(* IEC 61131-3 sources: PLC-IsaVODE/PLC-IsaVODE/samples/plc-programs (part 14) *)

(* ---- 100-RES_NTC.ST ---- *)
FUNCTION RES_NTC:REAL

	VAR_INPUT
		T :	REAL;
		RN :	REAL;
		B :	REAL;
	END_VAR

	RES_NTC := RN * EXP(B * (1.0 / (T+273.15) - 0.00335401643468053));

END_FUNCTION

PROGRAM program0

	VAR
		T :	REAL;
		RN :	REAL;
		B :	REAL;

		OUT :	REAL;
	END_VAR
		OUT := RES_NTC(T, RN, B);

END_PROGRAM

CONFIGURATION Config0

	RESOURCE Res0 ON PLC
		TASK task0(INTERVAL := T#20ms,PRIORITY := 0);
		PROGRAM instance0 WITH task0 : program0;
	END_RESOURCE

END_CONFIGURATION

(* ---- 101-WINDOW2.ST ---- *)
FUNCTION WINDOW2:BOOL
	VAR_INPUT
		LOW :	REAL;
		IN :	REAL;
		HIGH :	REAL;
	END_VAR
	window2 := (in <= high) AND (in >= low);
END_FUNCTION

PROGRAM program0
  	VAR
		LOW :	REAL;
		IN :	REAL;
		HIGH :	REAL;
		CEIL5_OUT : BOOL;
	END_VAR

  	CEIL5_OUT := window2(LOW, IN, HIGH);
END_PROGRAM

CONFIGURATION Config0
  	RESOURCE Res0 ON PLC
    	TASK task0(INTERVAL := T#20ms,PRIORITY := 0);
    	PROGRAM instance0 WITH task0 : program0;
  	END_RESOURCE
END_CONFIGURATION

(* ---- 102-F_LIN.ST ---- *)
FUNCTION F_LIN:REAL
	VAR_INPUT
		X :	REAL;
		A :	REAL;
		B :	REAL;
	END_VAR

	F_lin := A * X + B;
END_FUNCTION

PROGRAM program0
  VAR
    LocalVar0 : REAL;
	LocalVar1 : REAL;
	LocalVar2 : REAL;
	  LocalOUT  : REAL;
  END_VAR
  	LocalOUT := F_LIN(LocalVar0, LocalVar1, LocalVar2);
END_PROGRAM

CONFIGURATION Config0
  RESOURCE Res0 ON PLC
    TASK task0(INTERVAL := T#20ms,PRIORITY := 0);
    PROGRAM instance0 WITH task0 : program0;
  END_RESOURCE
END_CONFIGURATION

(* ---- 103-TN_SC_SHADOW_ATTR.ST ---- *)
FUNCTION TN_SC_SHADOW_ATTR:BYTE

	VAR_INPUT
		Iby_ATTR :	BYTE;
	END_VAR

	TN_SC_SHADOW_ATTR := ((Iby_ATTR AND BYTE#2#11110000) OR BYTE#2#00001000);

END_FUNCTION

PROGRAM program0
	VAR
		Iby_ATTR :	BYTE;
		CEIL5_OUT : BYTE;
	END_VAR

  	CEIL5_OUT := TN_SC_SHADOW_ATTR(Iby_ATTR);
END_PROGRAM

CONFIGURATION Config0

  RESOURCE Res0 ON PLC
    TASK task0(INTERVAL := T#20ms,PRIORITY := 0);
    PROGRAM instance0 WITH task0 : program0;
  END_RESOURCE
END_CONFIGURATION

(* ---- 104-DEC1.ST ---- *)
FUNCTION DEC1:INT

	VAR_INPUT
		X :	INT;
		N :	INT;
	END_VAR

	IF X = 0 THEN
		DEC1 := N - 1;
	ELSE
		DEC1 := X - 1;
	END_IF;

END_FUNCTION

PROGRAM program0
  VAR
    LocalVar0 : INT;
	LocalVar1 : INT;
	LocalOUT  : INT;
  END_VAR
  	LocalOUT := DEC1(LocalVar0, LocalVar1);
END_PROGRAM

CONFIGURATION Config0
  RESOURCE Res0 ON PLC
    TASK task0(INTERVAL := T#20ms,PRIORITY := 0);
    PROGRAM instance0 WITH task0 : program0;
  END_RESOURCE
END_CONFIGURATION

(* ---- 105-INC.ST ---- *)
FUNCTION INC:INT
	VAR_INPUT
		X :	INT;
		D :	INT;
		M :	INT;
	END_VAR

	inc := (X + D + M + 1) MOD (M + 1);
END_FUNCTION

PROGRAM program0
  VAR
    LocalVar0 : INT;
	LocalVar1 : INT;
	LocalVar2 : INT;
	LocalOUT  : INT;
  END_VAR
  	LocalOUT := INC(LocalVar0, LocalVar1,LocalVar2);
END_PROGRAM

CONFIGURATION Config0
  RESOURCE Res0 ON PLC
    TASK task0(INTERVAL := T#20ms,PRIORITY := 0);
    PROGRAM instance0 WITH task0 : program0;
  END_RESOURCE
END_CONFIGURATION

(* ---- 106-BIT_TOGGLE_B.ST ---- *)
FUNCTION BIT_TOGGLE_B:BYTE
	VAR_INPUT
		IN :	BYTE;
		POS :	INT;
	END_VAR

	BIT_TOGGLE_B := SHL(BYTE#1, POS) XOR IN;
END_FUNCTION

PROGRAM program0
  VAR
    LocalVar0 : BYTE;
    LocalVar1 : INT;
    CEIL5_OUT : BYTE;
  END_VAR

  CEIL5_OUT := BIT_TOGGLE_B(LocalVar0, LocalVar1);
END_PROGRAM

CONFIGURATION Config0

  RESOURCE Res0 ON PLC
    TASK task0(INTERVAL := T#20ms,PRIORITY := 0);
    PROGRAM instance0 WITH task0 : program0;
  END_RESOURCE
END_CONFIGURATION

(* ---- 107-BIT_TOGGLE_W.ST ---- *)
FUNCTION BIT_TOGGLE_W:WORD
	VAR_INPUT
		IN :	WORD;
		POS :	INT;
	END_VAR

	BIT_TOGGLE_W := SHL(WORD#1, POS) XOR IN;
END_FUNCTION

PROGRAM program0
  VAR
    LocalVar0 : WORD;
    LocalVar1 : INT;
    CEIL5_OUT : WORD;
  END_VAR

  CEIL5_OUT := BIT_TOGGLE_W(LocalVar0, LocalVar1);
END_PROGRAM

CONFIGURATION Config0

  RESOURCE Res0 ON PLC
    TASK task0(INTERVAL := T#20ms,PRIORITY := 0);
    PROGRAM instance0 WITH task0 : program0;
  END_RESOURCE
END_CONFIGURATION

(* ---- 108-RES_NI.ST ---- *)
FUNCTION RES_NI:REAL

	VAR_INPUT
		T :	REAL;
		R0 :	REAL;
	END_VAR

	VAR
		T2 :	REAL;
	END_VAR

	T2 := T*T;
	Res_NI := R0 + 0.5485*T + 0.665E-3*T2 + 2.805E-9*T2*T2;

END_FUNCTION

PROGRAM program0

	VAR
		T :	REAL;
		R0 :	REAL;

		OUT :	REAL;
	END_VAR
	OUT := RES_NI(T, R0);

END_PROGRAM

CONFIGURATION Config0

	RESOURCE Res0 ON PLC
		TASK task0(INTERVAL := T#20ms,PRIORITY := 0);
		PROGRAM instance0 WITH task0 : program0;
	END_RESOURCE

END_CONFIGURATION

(* ---- 109-TANK_VOL2.ST ---- *)
FUNCTION TANK_VOL2:REAL

	VAR_INPUT
		TR :	REAL;
		H :	REAL;
	END_VAR

	TANK_VOL2 := 3.14159265358979323846264338327950288 * H * H * (TR - H / 3.0);

END_FUNCTION

PROGRAM program0
  VAR
    TR :	REAL;
	H :	REAL;
    CEIL5_OUT : REAL;
  END_VAR

  CEIL5_OUT := TANK_VOL2(TR, H);
END_PROGRAM

CONFIGURATION Config0

  RESOURCE Res0 ON PLC
    TASK task0(INTERVAL := T#20ms,PRIORITY := 0);
    PROGRAM instance0 WITH task0 : program0;
  END_RESOURCE
END_CONFIGURATION

(* ---- 11-SWAP_BYTE.ST ---- *)
FUNCTION SWAP_BYTE:WORD

	VAR_INPUT
		IN :	WORD;
	END_VAR

	Swap_Byte := ROL(in,8);

END_FUNCTION

PROGRAM program0

	VAR
		IN :	WORD;
		CEIL5_OUT : WORD;
	END_VAR

	CEIL5_OUT := SWAP_BYTE(IN);

END_PROGRAM

CONFIGURATION Config0

	RESOURCE Res0 ON PLC
		TASK task0(INTERVAL := T#20ms,PRIORITY := 0);
		PROGRAM instance0 WITH task0 : program0;
	END_RESOURCE

END_CONFIGURATION

(* ---- 110-YEAR_END.ST ---- *)
FUNCTION YEAR_END:UDINT

	VAR_INPUT
		Y :	INT;
	END_VAR

	YEAR_END := DWORD_TO_UDINT(SHR(UDINT_TO_DWORD(INT_TO_UDINT(y) * UDINT#1461 - UDINT#2876712), 2)) * UDINT#86400;

END_FUNCTION

PROGRAM program0
  VAR
    Y : INT;
    CEIL5_OUT : UDINT;
  END_VAR

  CEIL5_OUT := YEAR_END(Y);
END_PROGRAM

CONFIGURATION Config0

  RESOURCE Res0 ON PLC
    TASK task0(INTERVAL := T#20ms,PRIORITY := 0);
    PROGRAM instance0 WITH task0 : program0;
  END_RESOURCE
END_CONFIGURATION

(* ---- 111-IP4_CHECK.ST ---- *)
FUNCTION IP4_CHECK:BOOL

	VAR_INPUT
		NIP :	DWORD;
		LIP :	DWORD;
		SM :	DWORD;
	END_VAR

	IP4_CHECK := (NIP AND sm) = (LIP AND SM);

END_FUNCTION

PROGRAM program0
	VAR
		NIP :	DWORD;
		LIP :	DWORD;
		SM :	DWORD;
		CEIL5_OUT : BOOL;
	END_VAR

  	CEIL5_OUT := IP4_CHECK(NIP, LIP, SM);
END_PROGRAM

CONFIGURATION Config0

  RESOURCE Res0 ON PLC
    TASK task0(INTERVAL := T#20ms,PRIORITY := 0);
    PROGRAM instance0 WITH task0 : program0;
  END_RESOURCE
END_CONFIGURATION

(* ---- 112-ELLIPSE_A.ST ---- *)
FUNCTION ELLIPSE_A:REAL
	VAR_INPUT
		R1 :	REAL;
		R2 :	REAL;
	END_VAR

	ellipse_A := 3.14159265358979323846264338327950288 * R1 * R2;

END_FUNCTION

PROGRAM program0
  VAR
    LocalVar0 : REAL;
	LocalVar1 : REAL;
	  LocalOUT  : REAL;
  END_VAR
  	LocalOUT := ELLIPSE_A(LocalVar0, LocalVar1);
END_PROGRAM

CONFIGURATION Config0
  RESOURCE Res0 ON PLC
    TASK task0(INTERVAL := T#20ms,PRIORITY := 0);
    PROGRAM instance0 WITH task0 : program0;
  END_RESOURCE
END_CONFIGURATION

(* ---- 113-F_POWER.ST ---- *)
FUNCTION F_POWER:REAL
	VAR_INPUT
		A :	REAL;
		X :	REAL;
		N :	REAL;
	END_VAR

	f_power := a * EXPT(X,N);
END_FUNCTION

PROGRAM program0
  VAR
    LocalVar0 : REAL;
	LocalVar1 : REAL;
	LocalVar2 : REAL;
	  LocalOUT  : REAL;
  END_VAR
  	LocalOUT := F_POWER(LocalVar0, LocalVar1, LocalVar2);
END_PROGRAM

CONFIGURATION Config0
  RESOURCE Res0 ON PLC
    TASK task0(INTERVAL := T#20ms,PRIORITY := 0);
    PROGRAM instance0 WITH task0 : program0;
  END_RESOURCE
END_CONFIGURATION

(* ---- 114-TANH.ST ---- *)
FUNCTION TANH:REAL

	VAR_INPUT
		X :	REAL;
	END_VAR

	IF X > 20.0 THEN
		TANH := 1.0;
	ELSIF X < -20.0 THEN
		TANH := -1.0;
	ELSE
		TANH := 1.0 - 2.0 / (EXP(2.0 * x) + 1.0);
	END_IF;

END_FUNCTION

PROGRAM program0

	VAR
		X :	REAL;
		CEIL5_OUT : REAL;
	END_VAR

	CEIL5_OUT := TANH(X);

END_PROGRAM

CONFIGURATION Config0

	RESOURCE Res0 ON PLC
		TASK task0(INTERVAL := T#20ms,PRIORITY := 0);
		PROGRAM instance0 WITH task0 : program0;
	END_RESOURCE

END_CONFIGURATION

(* ---- 115-BIT_TOGGLE_DW.ST ---- *)
FUNCTION BIT_TOGGLE_DW:DWORD
	VAR_INPUT
		IN :	DWORD;
		POS :	INT;
	END_VAR

	BIT_TOGGLE_DW := SHL(DWORD#1, POS) XOR IN;

END_FUNCTION

PROGRAM program0
  VAR
    LocalVar0 : DWORD;
    LocalVar1 : INT;
    CEIL5_OUT : DWORD;
  END_VAR

  CEIL5_OUT := BIT_TOGGLE_DW(LocalVar0, LocalVar1);
END_PROGRAM

CONFIGURATION Config0

  RESOURCE Res0 ON PLC
    TASK task0(INTERVAL := T#20ms,PRIORITY := 0);
    PROGRAM instance0 WITH task0 : program0;
  END_RESOURCE
END_CONFIGURATION

(* ---- 116-SIGMOID.ST ---- *)
FUNCTION SIGMOID:REAL

	VAR_INPUT
		X :	REAL;
	END_VAR

	IF X > 20.0 THEN
		SIGMOID := 1.0;
	ELSIF x < -85.0 THEN
		SIGMOID := 0.0;
	ELSE
		SIGMOID := 1.0 / (1.0 + EXP(-X));
	END_IF;

END_FUNCTION

PROGRAM program0

	VAR
		X :	REAL;
		CEIL5_OUT : REAL;
	END_VAR

	CEIL5_OUT := SIGMOID(X);

END_PROGRAM

CONFIGURATION Config0

	RESOURCE Res0 ON PLC
		TASK task0(INTERVAL := T#20ms,PRIORITY := 0);
		PROGRAM instance0 WITH task0 : program0;
	END_RESOURCE

END_CONFIGURATION

(* ---- 117-LEAP_OF_DATE.ST ---- *)
FUNCTION LEAP_OF_DATE:BOOL

	VAR_INPUT
		IDATE :	UDINT;
	END_VAR

	LEAP_OF_DATE := SHL(UDINT_TO_DWORD((idate + UDINT#43200) / UDINT#31557600), 30) = DWORD#16#80000000;

END_FUNCTION

PROGRAM program0
  VAR
    LocalVar0 : UDINT;
	LocalOUT  : BOOL;
  END_VAR
  	LocalOUT := LEAP_OF_DATE(LocalVar0);
END_PROGRAM

CONFIGURATION Config0
  RESOURCE Res0 ON PLC
    TASK task0(INTERVAL := T#20ms,PRIORITY := 0);
    PROGRAM instance0 WITH task0 : program0;
  END_RESOURCE
END_CONFIGURATION

(* ---- 118-DIFFER.ST ---- *)
FUNCTION DIFFER:BOOL
	VAR_INPUT
		IN1 :	REAL;
		IN2 :	REAL;
		X :	REAL;
	END_VAR

	DIFFER := ABS(in1 - in2) > X;
END_FUNCTION

PROGRAM program0
  VAR
    LocalVar0 : REAL;
	LocalVar1 : REAL;
	LocalVar2 : REAL;
	LocalOUT  : BOOL;
  END_VAR
  	LocalOUT := DIFFER(LocalVar0, LocalVar1, LocalVar2);
END_PROGRAM

CONFIGURATION Config0
  RESOURCE Res0 ON PLC
    TASK task0(INTERVAL := T#20ms,PRIORITY := 0);
    PROGRAM instance0 WITH task0 : program0;
  END_RESOURCE
END_CONFIGURATION

(* ---- 119-DEAD_ZONE.ST ---- *)
FUNCTION DEAD_ZONE:REAL

	VAR_INPUT
		X :	REAL;
		L :	REAL;
	END_VAR

	IF ABS(x) > L THEN
		dead_zone := X;
	ELSE
		DEAD_ZONE := 0.0;
	END_IF;

END_FUNCTION

PROGRAM program0
  VAR
    LocalVar0 : REAL;
	LocalVar1 : REAL;
	LocalOUT  : REAL;
  END_VAR
  	LocalOUT := DEAD_ZONE(LocalVar0, LocalVar1);
END_PROGRAM

CONFIGURATION Config0
  RESOURCE Res0 ON PLC
    TASK task0(INTERVAL := T#20ms,PRIORITY := 0);
    PROGRAM instance0 WITH task0 : program0;
  END_RESOURCE
END_CONFIGURATION

(* ---- 12-ISC_CTRL.ST ---- *)
FUNCTION ISC_CTRL:BOOL

	VAR_INPUT
		IN :	BYTE;
	END_VAR

	ISC_CTRL := IN < BYTE#32 OR IN = BYTE#127;

END_FUNCTION

PROGRAM program0
	VAR
		IN : BYTE;
		OUT : BOOL;
	END_VAR

	OUT := ISC_CTRL(IN);
END_PROGRAM

CONFIGURATION Config0

	RESOURCE Res0 ON PLC
		TASK task0(INTERVAL := T#20ms,PRIORITY := 0);
		PROGRAM instance0 WITH task0 : program0;
	END_RESOURCE

END_CONFIGURATION

(* ---- 120-SQRTN.ST ---- *)
FUNCTION SQRTN:REAL

	VAR_INPUT
		X :	REAL;
		N :	INT;
	END_VAR

	IF N > 0 THEN
		SQRTN := EXP(LN(x) / INT_TO_REAL(n));
	ELSE
		SQRTN := 0.0;
	END_IF;

END_FUNCTION

PROGRAM program0
	VAR
		LocalVar0 : REAL;
		LocalVar1 : INT;
		LocalOUT  : REAL;
	END_VAR

 	LocalOUT := SQRTN(LocalVar0, LocalVar1);

END_PROGRAM

CONFIGURATION Config0

	RESOURCE Res0 ON PLC
		TASK task0(INTERVAL := T#20ms,PRIORITY := 0);
		PROGRAM instance0 WITH task0 : program0;
	END_RESOURCE

END_CONFIGURATION

(* ---- 122-DWORD_OF_WORD.ST ---- *)
FUNCTION DWORD_OF_WORD:DWORD

	VAR_INPUT
		W1 :	WORD;
		W0 :	WORD;
	END_VAR

	DWORD_OF_WORD := SHL(WORD_TO_DWORD(W1),16) OR WORD_TO_DWORD(W0);

END_FUNCTION

PROGRAM program0
  VAR
    LocalVar0 : WORD;
	LocalVar1 : WORD;
	LocalOUT  : DWORD;
  END_VAR
  	LocalOUT := DWORD_OF_WORD(LocalVar0, LocalVar1);
END_PROGRAM

CONFIGURATION Config0
  RESOURCE Res0 ON PLC
    TASK task0(INTERVAL := T#20ms,PRIORITY := 0);
    PROGRAM instance0 WITH task0 : program0;
  END_RESOURCE
END_CONFIGURATION

(* ---- 123-WCT.ST ---- *)
FUNCTION WCT:REAL

	VAR_INPUT
		T :	REAL;
		V :	REAL;
	END_VAR

	IF V < 5.0 OR T > 10.0 THEN
		WCT := T;
	ELSE
		WCT := 13.12 + 0.6215 * T +(0.3965 * T - 11.37) * EXP(LN(v) * 0.16);
	END_IF;

END_FUNCTION

PROGRAM program0
	VAR
		T :	REAL;
		V :	REAL;
		CEIL5_OUT : REAL;
	END_VAR

  	CEIL5_OUT := WCT(T, V);
END_PROGRAM

CONFIGURATION Config0

  RESOURCE Res0 ON PLC
    TASK task0(INTERVAL := T#20ms,PRIORITY := 0);
    PROGRAM instance0 WITH task0 : program0;
  END_RESOURCE
END_CONFIGURATION

(* ---- 124-TEMP_NTC.ST ---- *)
FUNCTION TEMP_NTC:REAL

VAR_INPUT
	RES :	REAL;
	RN :	REAL;
	B :	REAL;
END_VAR

IF res > 0.0 THEN
	TEMP_NTC := B * 298.15 / (B + LN(RES / RN) * 298.15) -273.15;
END_IF;

END_FUNCTION

PROGRAM program0
  	VAR
		RES :	REAL;
		RN :	REAL;
		B :	REAL;
    	CEIL5_OUT : REAL;
  	END_VAR

  	CEIL5_OUT := TEMP_NTC(RES, RN, B);
END_PROGRAM

CONFIGURATION Config0
	RESOURCE Res0 ON PLC
		TASK task0(INTERVAL := T#20ms,PRIORITY := 0);
		PROGRAM instance0 WITH task0 : program0;
	END_RESOURCE
END_CONFIGURATION

(* ---- 125-SCALE.ST ---- *)
FUNCTION SCALE:REAL

	VAR_INPUT
		X :	REAL;
		K :	REAL;
		O :	REAL;
		MX :	REAL;
		MN :	REAL;
	END_VAR

	SCALE := LIMIT(MN, X * K + O, MX);

END_FUNCTION

PROGRAM program0
  VAR
    X :	REAL;
	K :	REAL;
	O :	REAL;
	MX :	REAL;
	MN :	REAL;
    CEIL5_OUT : REAL;
  END_VAR

  CEIL5_OUT := SCALE(X, K, O, MX, MN);
END_PROGRAM

CONFIGURATION Config0

  RESOURCE Res0 ON PLC
    TASK task0(INTERVAL := T#20ms,PRIORITY := 0);
    PROGRAM instance0 WITH task0 : program0;
  END_RESOURCE
END_CONFIGURATION

(* ---- 126-_MOD_INT.ST ---- *)
FUNCTION _MOD_INT:INT
  VAR_INPUT
    IN :	INT;
    DIVISOR :	INT;
  END_VAR

  IF IN = 0 THEN
    _MOD_INT := 0;
  ELSE
    _MOD_INT := IN MOD DIVISOR;
  END_IF;
END_FUNCTION

PROGRAM program0
  VAR
    LocalVar0 : INT;
    LocalVar1 : INT;
	  LocalOUT  : INT;
  END_VAR

  LocalOUT := _MOD_INT(LocalVar0, LocalVar1);
END_PROGRAM

CONFIGURATION Config0
  RESOURCE Res0 ON PLC
    TASK task0(INTERVAL := T#20ms,PRIORITY := 0);
    PROGRAM instance0 WITH task0 : program0;
  END_RESOURCE
END_CONFIGURATION

(* ---- 127-INC2.ST ---- *)
FUNCTION INC2:INT

	VAR_INPUT
		X :	INT;
		D :	INT;
		L :	INT;
		U :	INT;
	END_VAR

	VAR
		tmp :	INT;
	END_VAR

	tmp := U - L + 1;
	INC2 := (X + D - L + tmp) MOD tmp + L;

END_FUNCTION

PROGRAM program0
	VAR
		X :	INT;
		D :	INT;
		L :	INT;
		U :	INT;
		CEIL5_OUT : INT;
	END_VAR

  	CEIL5_OUT := INC2(X, D, L, U);
END_PROGRAM

CONFIGURATION Config0

	RESOURCE Res0 ON PLC
		TASK task0(INTERVAL := T#20ms,PRIORITY := 0);
		PROGRAM instance0 WITH task0 : program0;
	END_RESOURCE

END_CONFIGURATION

(* ---- 128-TEMP_SI.ST ---- *)
FUNCTION TEMP_SI:REAL
	VAR_INPUT
		RES :	REAL;
		VAR_RS:	REAL;
		TS :	REAL;
	END_VAR

	TEMP_SI := (-7.64E-3 + SQRT(RES/VAR_RS* 6.64E-5 - 0.803E-5)) * 30120.48193 + TS;

END_FUNCTION

PROGRAM program0
  	VAR
		RES :	REAL;
		VAR_RS:	REAL;
		TS :	REAL;
    	CEIL5_OUT : REAL;
  	END_VAR

  	CEIL5_OUT := TEMP_SI(RES, VAR_RS, TS);
END_PROGRAM

CONFIGURATION Config0
	RESOURCE Res0 ON PLC
		TASK task0(INTERVAL := T#20ms,PRIORITY := 0);
		PROGRAM instance0 WITH task0 : program0;
	END_RESOURCE
END_CONFIGURATION

(* ---- 129-CAUCHYCD.ST ---- *)
FUNCTION CAUCHYCD:REAL
	VAR_INPUT
		X :	REAL;
		T :	REAL;
		U :	REAL;
	END_VAR

	CAUCHYCD := 0.5 + 0.318309886183791 * ATAN((X - T) / U);
END_FUNCTION

PROGRAM program0
  VAR
    LocalVar0 : REAL;
	LocalVar1 : REAL;
	LocalVar2 : REAL;
	LocalOUT  : REAL;
  END_VAR
	LocalOUT := CAUCHYCD(LocalVar0, LocalVar1, LocalVar2);
END_PROGRAM

CONFIGURATION Config0
  RESOURCE Res0 ON PLC
    TASK task0(INTERVAL := T#20ms,PRIORITY := 0);
    PROGRAM instance0 WITH task0 : program0;
  END_RESOURCE
END_CONFIGURATION

(* ---- 13-KMH_TO_MS.ST ---- *)
FUNCTION KMH_TO_MS:REAL

	VAR_INPUT
		KMH :	REAL;
	END_VAR

	KMH_TO_MS := kmh * 0.2777777777777;

END_FUNCTION

PROGRAM program0
	VAR
		KMH : REAL;
		OUT : REAL;
	END_VAR

	OUT := KMH_TO_MS(KMH);
END_PROGRAM

CONFIGURATION Config0

	RESOURCE Res0 ON PLC
		TASK task0(INTERVAL := T#20ms,PRIORITY := 0);
		PROGRAM instance0 WITH task0 : program0;
	END_RESOURCE

END_CONFIGURATION

(* ---- 130-FLOOR.ST ---- *)
FUNCTION FLOOR : INT
  VAR_INPUT
    x : REAL;
  END_VAR

  FLOOR := REAL_TO_INT(X);
  IF INT_TO_REAL(FLOOR) > X THEN
  	floor := floor - 1;
  END_IF;
  (* from OSCAT library; www.oscat.de  *)
END_FUNCTION

PROGRAM program0
  VAR
    LocalVar0 : REAL;
    CEIL5_OUT : INT;
  END_VAR

  CEIL5_OUT := FLOOR(LocalVar0);
END_PROGRAM

CONFIGURATION Config0

  RESOURCE Res0 ON PLC
    TASK task0(INTERVAL := T#20ms,PRIORITY := 0);
    PROGRAM instance0 WITH task0 : program0;
  END_RESOURCE
END_CONFIGURATION

(* ---- 131-GAMMA.ST ---- *)
FUNCTION GAMMA:REAL
	VAR_INPUT
		X :	REAL;
	END_VAR

	IF x > 0.0 THEN
		GAMMA := SQRT(6.28318530717958647692528676655900576 / X) * EXPT(0.367879441171442 * (x + 1.0 / (12.0 * x - 0.1 / X)), X);
	END_IF;
END_FUNCTION

PROGRAM program0
  VAR
    LocalVar0 : REAL;
    LocalOUT  : REAL;
  END_VAR

  LocalOUT := GAMMA(LocalVar0);
END_PROGRAM

CONFIGURATION Config0
  RESOURCE Res0 ON PLC
    TASK task0(INTERVAL := T#20ms,PRIORITY := 0);
    PROGRAM instance0 WITH task0 : program0;
  END_RESOURCE
END_CONFIGURATION

(* ---- 132-REFRACTION.ST ---- *)
FUNCTION REFRACTION:REAL

	VAR_INPUT
		ELEV :	REAL;
	END_VAR

	VAR
		tmp :	REAL;
	END_VAR

	tmp := LIMIT(-1.9, elev, 80.0);
	REFRACTION := 0.0174532925199433 / TAN(0.0174532925199433 * (tmp + 10.3 / (tmp + 5.11)));

END_FUNCTION

PROGRAM program0

	VAR
		ELEV :	REAL;

		OUT :	REAL;
	END_VAR
	OUT := REFRACTION(ELEV);

END_PROGRAM

CONFIGURATION Config0

	RESOURCE Res0 ON PLC
		TASK task0(INTERVAL := T#20ms,PRIORITY := 0);
		PROGRAM instance0 WITH task0 : program0;
	END_RESOURCE

END_CONFIGURATION

(* ---- 133-GEO_TO_DEG.ST ---- *)
FUNCTION GEO_TO_DEG:REAL

	VAR_INPUT
		D :	INT;
		M :	INT;
		SEC :	REAL;
	END_VAR

	GEO_TO_DEG := INT_TO_REAL(D) + INT_TO_REAL(M) * 0.016666666666667 + sec * 0.00027777777777778;

END_FUNCTION

PROGRAM program0
  VAR
    D :	INT;
	M :	INT;
	SEC :	REAL;
    LocalOUT  : REAL;
  END_VAR

  LocalOUT := GEO_TO_DEG(D, M, SEC);
END_PROGRAM

CONFIGURATION Config0
  RESOURCE Res0 ON PLC
    TASK task0(INTERVAL := T#20ms,PRIORITY := 0);
    PROGRAM instance0 WITH task0 : program0;
  END_RESOURCE
END_CONFIGURATION

(* ---- 134-GRAY_TO_BYTE.ST ---- *)
FUNCTION GRAY_TO_BYTE:BYTE

	VAR_INPUT
		IN :	BYTE;
	END_VAR

	GRAY_TO_BYTE := SHR(IN,4) XOR IN;
	GRAY_TO_BYTE := SHR(GRAY_TO_BYTE,2) XOR GRAY_TO_BYTE;
	GRAY_TO_BYTE := SHR(GRAY_TO_BYTE,1) XOR GRAY_TO_BYTE;

END_FUNCTION

PROGRAM program0
  VAR
   	IN :	BYTE;
    LocalOUT  : BYTE;
  END_VAR

  LocalOUT := GRAY_TO_BYTE(IN);
END_PROGRAM

CONFIGURATION Config0
  RESOURCE Res0 ON PLC
    TASK task0(INTERVAL := T#20ms,PRIORITY := 0);
    PROGRAM instance0 WITH task0 : program0;
  END_RESOURCE
END_CONFIGURATION

(* ---- 135-RES_SI.ST ---- *)
FUNCTION RES_SI:REAL

	VAR_INPUT
		T :	REAL;
		_RS :	REAL;
		TS :	REAL;
	END_VAR

	VAR
		TX :	REAL;
	END_VAR

	TX := T - TS;
	RES_SI := _RS * ( 1.0 + 7.64E-3 * TX + 1.66E-5 * TX * TX);

END_FUNCTION

PROGRAM program0

	VAR
		T :	REAL;
		_RS :	REAL;
		TS :	REAL;

		OUT :	REAL;
	END_VAR
		OUT := RES_SI(T, _RS, TS);

END_PROGRAM

CONFIGURATION Config0

	RESOURCE Res0 ON PLC
		TASK task0(INTERVAL := T#20ms,PRIORITY := 0);
		PROGRAM instance0 WITH task0 : program0;
	END_RESOURCE

END_CONFIGURATION

(* ---- 136-SDD.ST ---- *)
FUNCTION SDD:REAL

	VAR_INPUT
		T :	REAL;
		ICE :	BOOL;
	END_VAR

	IF ice THEN
		SDD := 611.153 * EXP(22.4433 * T / (272.186 + T));
	ELSE
		SDD := 611.213 * EXP(17.5043 * T / (241.2 + T));
	END_IF;

END_FUNCTION

PROGRAM program0
  VAR
    T :	REAL;
	ICE :	BOOL;
    CEIL5_OUT : REAL;
  END_VAR

  CEIL5_OUT := SDD(T, ICE);
END_PROGRAM

CONFIGURATION Config0

  RESOURCE Res0 ON PLC
    TASK task0(INTERVAL := T#20ms,PRIORITY := 0);
    PROGRAM instance0 WITH task0 : program0;
  END_RESOURCE
END_CONFIGURATION

(* ---- 137-SGN.ST ---- *)
FUNCTION SGN : INT
  VAR_INPUT
    x : REAL;
  END_VAR

  IF X > 0.0 THEN
  	sgn := 1;
  ELSIF X < 0.0 THEN
  	sgn := -1;
  ELSE
  	sgn := 0;
  END_IF;
END_FUNCTION

PROGRAM program0
  VAR
    LocalVar0 : REAL;
    LocalVar1 : INT;
    CEIL5_OUT : INT;
  END_VAR

  CEIL5_OUT := SGN(LocalVar0);
  LocalVar1 := CEIL5_OUT;
END_PROGRAM

CONFIGURATION Config0

  RESOURCE Res0 ON PLC
    TASK task0(INTERVAL := T#20ms,PRIORITY := 0);
    PROGRAM instance0 WITH task0 : program0;
  END_RESOURCE
END_CONFIGURATION

(* ---- 138-ELLIPSE_C.ST ---- *)
FUNCTION ELLIPSE_C:REAL

VAR_INPUT
	R1 :	REAL;
	R2 :	REAL;
END_VAR

ELLIPSE_C := 3.14159265358979323846264338327950288 * (3.0 * (R1+R2) - SQRT((3.0 * r1 + R2) * (3.0 * r2 + r1)));

END_FUNCTION

PROGRAM program0
  VAR
    LocalVar0 : REAL;
	LocalVar1 : REAL;
	  LocalOUT  : REAL;
  END_VAR
  	LocalOUT := ELLIPSE_C(LocalVar0, LocalVar1);
END_PROGRAM

CONFIGURATION Config0
  RESOURCE Res0 ON PLC
    TASK task0(INTERVAL := T#20ms,PRIORITY := 0);
    PROGRAM instance0 WITH task0 : program0;
  END_RESOURCE
END_CONFIGURATION

(* ---- 139-F_QUAD.ST ---- *)
FUNCTION F_QUAD:REAL

	VAR_INPUT
		X :	REAL;
		A :	REAL;
		B :	REAL;
		C :	REAL;
	END_VAR

	F_QUAD :=  (A * X + B) * X + C;

END_FUNCTION

PROGRAM program0
  VAR
    LocalVar0 : REAL;
	LocalVar1 : REAL;
	LocalVar2 : REAL;
	LocalVar3 : REAL;
	LocalOUT  : REAL;
  END_VAR
  	LocalOUT := F_QUAD(LocalVar0, LocalVar1, LocalVar2, LocalVar3);
END_PROGRAM

CONFIGURATION Config0
  RESOURCE Res0 ON PLC
    TASK task0(INTERVAL := T#20ms,PRIORITY := 0);
    PROGRAM instance0 WITH task0 : program0;
  END_RESOURCE
END_CONFIGURATION

(* ---- 14-GOLD.ST ---- *)
FUNCTION GOLD:REAL

	VAR_INPUT
		X :	REAL;
	END_VAR

	GOLD := (X + SQRT(X*X + 4.0)) * 0.5;

END_FUNCTION

PROGRAM program0
  VAR
   	X :	REAL;
    LocalOUT  : REAL;
  END_VAR

  LocalOUT := GOLD(X);
END_PROGRAM

CONFIGURATION Config0
  RESOURCE Res0 ON PLC
    TASK task0(INTERVAL := T#20ms,PRIORITY := 0);
    PROGRAM instance0 WITH task0 : program0;
  END_RESOURCE
END_CONFIGURATION

(* ---- 140-SDD_NH3.ST ---- *)
FUNCTION SDD_NH3:REAL

	VAR_INPUT
		T :	REAL;
	END_VAR

	IF T < -33.65 THEN
		SDD_NH3 := EXP(7.3396511649 - ( 1166.7498002 / ( T + 192.37 )));
	ELSE
		SDD_NH3 := EXP(11.210964456 - ( 2564.9140075 / ( T + 262.741 )));
	END_IF;

END_FUNCTION

PROGRAM program0
  VAR
    T :	REAL;
    CEIL5_OUT : REAL;
  END_VAR

  CEIL5_OUT := SDD_NH3(T);
END_PROGRAM

CONFIGURATION Config0

  RESOURCE Res0 ON PLC
    TASK task0(INTERVAL := T#20ms,PRIORITY := 0);
    PROGRAM instance0 WITH task0 : program0;
  END_RESOURCE
END_CONFIGURATION

(* ---- 142-DEAD_BAND.ST ---- *)
FUNCTION DEAD_BAND:REAL

	VAR_INPUT
		X :	REAL;
		L :	REAL;
	END_VAR

	IF X > L THEN
		DEAD_BAND := X - L;
	ELSIF X < -L THEN
		DEAD_BAND := X + L;
	ELSE
		DEAD_BAND := 0.0;
	END_IF;

END_FUNCTION

PROGRAM program0
  VAR
    LocalVar0 : REAL;
	LocalVar1 : REAL;
	LocalOUT  : REAL;
  END_VAR
  	LocalOUT := DEAD_BAND(LocalVar0, LocalVar1);
END_PROGRAM

CONFIGURATION Config0
  RESOURCE Res0 ON PLC
    TASK task0(INTERVAL := T#20ms,PRIORITY := 0);
    PROGRAM instance0 WITH task0 : program0;
  END_RESOURCE
END_CONFIGURATION

(* ---- 143-REVERSE.ST ---- *)
FUNCTION REVERSE:BYTE
VAR_INPUT
	IN :	BYTE;
END_VAR

reverse := SHL(in,7) OR SHR(in,7) OR (ROR(in,3) AND BYTE#2#01000100) OR (ROL(in,3) AND BYTE#2#00100010)
	OR (SHL(in,1) AND BYTE#2#00010000) OR (SHR(in,1) AND BYTE#2#00001000);

END_FUNCTION

PROGRAM program0
  VAR
    LocalVar0 : BYTE;
	LocalOUT  : BYTE;
  END_VAR
  	LocalOUT := REVERSE(LocalVar0);
END_PROGRAM

CONFIGURATION Config0
  RESOURCE Res0 ON PLC
    TASK task0(INTERVAL := T#20ms,PRIORITY := 0);
    PROGRAM instance0 WITH task0 : program0;
  END_RESOURCE
END_CONFIGURATION

(* ---- 144-BIT_OF_DWORD.ST ---- *)
FUNCTION BIT_OF_DWORD : BOOL
  VAR_INPUT
    IN : DWORD;
    N : INT;
  END_VAR

  BIT_OF_DWORD := (SHR(in,N) AND 16#00000001) > 0;
END_FUNCTION

PROGRAM program0
  VAR
    LocalVar0 : DWORD;
    LocalVar2 : INT;
    LocalVar1 : BOOL;
    CEIL5_OUT : BOOL;
  END_VAR

  CEIL5_OUT := BIT_OF_DWORD(LocalVar0, LocalVar2);
  LocalVar1 := CEIL5_OUT;
END_PROGRAM

CONFIGURATION Config0

  RESOURCE Res0 ON PLC
    TASK task0(INTERVAL := T#20ms,PRIORITY := 0);
    PROGRAM instance0 WITH task0 : program0;
  END_RESOURCE
END_CONFIGURATION

(* ---- 145-IS_URLCHR.ST ---- *)
FUNCTION IS_URLCHR:BOOL

	VAR_INPUT
		IN :	BYTE;
	END_VAR

	IS_URLCHR := ((IN>BYTE#47) AND (IN<BYTE#58)) OR ((IN>BYTE#64) AND (IN<BYTE#91)) OR ((IN>BYTE#96) AND (IN<BYTE#123)) OR (in=BYTE#126) OR (in=BYTE#95) OR (in=BYTE#45) OR (in=BYTE#46);

END_FUNCTION

PROGRAM program0
	VAR
		IN :	BYTE;
		CEIL5_OUT : BOOL;
	END_VAR

  	CEIL5_OUT := IS_URLCHR(IN);
END_PROGRAM

CONFIGURATION Config0

  RESOURCE Res0 ON PLC
    TASK task0(INTERVAL := T#20ms,PRIORITY := 0);
    PROGRAM instance0 WITH task0 : program0;
  END_RESOURCE
END_CONFIGURATION

(* ---- 146-GDF.ST ---- *)
FUNCTION GDF:REAL

	VAR_INPUT
		X :	REAL;
	END_VAR

	IF X = 0.0 THEN
		GDF := 0.0;
	ELSIF X > 15.0 THEN
		GDF := 1.5707963267949;
	ELSIF X < -15.0 THEN
		GDF := -1.5707963267949;
	ELSE
		GDF := ATAN(EXP(X)) * 2.0 - 1.5707963267949;
	END_IF;

END_FUNCTION

PROGRAM program0
  VAR
    X :	REAL;
    LocalOUT  : REAL;
  END_VAR

  LocalOUT := GDF(X);
END_PROGRAM

CONFIGURATION Config0
  RESOURCE Res0 ON PLC
    TASK task0(INTERVAL := T#20ms,PRIORITY := 0);
    PROGRAM instance0 WITH task0 : program0;
  END_RESOURCE
END_CONFIGURATION

(* ---- 147-SDT_NH3.ST ---- *)
FUNCTION SDT_NH3:REAL

	VAR_INPUT
		P :	REAL;
	END_VAR

	IF P < 1.0E-3 THEN
		SDT_NH3 := -110.0;
	ELSIF P < 1.0 THEN
		SDT_NH3 := 506.713 / (3.18757 - LOG(P)) - 192.37 ;
	ELSE
		SDT_NH3 := 1113.928 / (4.86886 - LOG(P)) - 262.71 ;
	END_IF;

END_FUNCTION

PROGRAM program0
  VAR
    P :	REAL;
    CEIL5_OUT : REAL;
  END_VAR

  CEIL5_OUT := SDT_NH3(P);
END_PROGRAM

CONFIGURATION Config0

  RESOURCE Res0 ON PLC
    TASK task0(INTERVAL := T#20ms,PRIORITY := 0);
    PROGRAM instance0 WITH task0 : program0;
  END_RESOURCE
END_CONFIGURATION

(* ---- 148-PT_TO_F.ST ---- *)
FUNCTION _DWORD_TO_REAL:REAL
	VAR_INPUT
		IN :	DWORD;
	END_VAR

	_DWORD_TO_REAL := UDINT_TO_REAL(DWORD_TO_UDINT(IN));

END_FUNCTION

FUNCTION PT_TO_F:REAL

	VAR_INPUT
		PT :	TIME;
	END_VAR

	PT_TO_F := 1000.0 / _DWORD_TO_REAL(TIME_TO_DWORD(PT));

END_FUNCTION

PROGRAM program0
  VAR
    PT : TIME;
    OUT : REAL;
  END_VAR

  OUT := PT_TO_F(PT);
END_PROGRAM

CONFIGURATION Config0

  RESOURCE Res0 ON PLC
    TASK task0(INTERVAL := T#20ms,PRIORITY := 0);
    PROGRAM instance0 WITH task0 : program0;
  END_RESOURCE
END_CONFIGURATION

(* ---- 15-DATE_TO_DT.ST ---- *)
FUNCTION DATE_TO_DT:UDINT
	VAR_INPUT
		IN :	UDINT;
	END_VAR
	DATE_TO_DT := IN;
END_FUNCTION

PROGRAM program0
  VAR
    LocalVar0 : UDINT;
	LocalOUT  : UDINT;
  END_VAR
  	LocalOUT := DATE_TO_DT(LocalVar0);
END_PROGRAM

CONFIGURATION Config0
  RESOURCE Res0 ON PLC
    TASK task0(INTERVAL := T#20ms,PRIORITY := 0);
    PROGRAM instance0 WITH task0 : program0;
  END_RESOURCE
END_CONFIGURATION

(* ---- 150-SIGN_I.ST ---- *)
FUNCTION BIT_OF_DWORD : BOOL

	VAR_INPUT
		IN : DWORD;
		N : INT;
	END_VAR

	BIT_OF_DWORD := (SHR(in,N) AND 16#00000001) > 0;

END_FUNCTION

FUNCTION SIGN_I:BOOL

	VAR_INPUT
		IN :	DINT;
	END_VAR

	sign_I := BIT_OF_DWORD(DINT_TO_DWORD(in),31);

END_FUNCTION

PROGRAM program0

	VAR
		IN :	DINT;
		CEIL5_OUT : BOOL;
	END_VAR

	CEIL5_OUT := SIGN_I(IN);

END_PROGRAM

CONFIGURATION Config0

	RESOURCE Res0 ON PLC
		TASK task0(INTERVAL := T#20ms,PRIORITY := 0);
		PROGRAM instance0 WITH task0 : program0;
	END_RESOURCE

END_CONFIGURATION

(* ---- 153-BAND_B.ST ---- *)
FUNCTION BAND_B:BYTE
	VAR_INPUT
		X :	BYTE;
		B :	BYTE;
	END_VAR

	IF X < B THEN
		BAND_B := BYTE#0;
	ELSIF X > USINT_TO_BYTE(USINT#255 - BYTE_TO_USINT(B)) THEN
		BAND_B := BYTE#255;
	ELSE
		BAND_B := X;
	END_IF;
END_FUNCTION
PROGRAM program0
  VAR
    LocalVar0 : BYTE;
	LocalVar1 : BYTE;
    LocalOUT  : BYTE;
  END_VAR

  LocalOUT := BAND_B(LocalVar0, LocalVar1);
END_PROGRAM

CONFIGURATION Config0
  RESOURCE Res0 ON PLC
    TASK task0(INTERVAL := T#20ms,PRIORITY := 0);
    PROGRAM instance0 WITH task0 : program0;
  END_RESOURCE
END_CONFIGURATION

(* ---- 154-CAUCHY.ST ---- *)
FUNCTION CAUCHY:REAL
	VAR_INPUT
		X :	REAL;
		T :	REAL;
		U :	REAL;
	END_VAR

	VAR
		tmp :	REAL;
	END_VAR

	tmp := x - t;
	CAUCHY := 0.318309886183791 * U / (U*U + tmp*tmp);
END_FUNCTION

PROGRAM program0
  VAR
    LocalVar0 : REAL;
    LocalVar1 : REAL;
	LocalVar2 : REAL;
    CEIL5_OUT : REAL;
  END_VAR

  CEIL5_OUT := CAUCHY(LocalVar0, LocalVar1, LocalVar2);
END_PROGRAM

CONFIGURATION Config0

  RESOURCE Res0 ON PLC
    TASK task0(INTERVAL := T#20ms,PRIORITY := 0);
    PROGRAM instance0 WITH task0 : program0;
  END_RESOURCE
END_CONFIGURATION

(* ---- 155-TN_SC_XY2_ERROR.ST ---- *)
FUNCTION TN_SC_XY2_ERROR:BOOL

	VAR_INPUT
		X1 :	INT;
		Y1 :	INT;
		X2 :	INT;
		Y2 :	INT;
	END_VAR

	TN_SC_XY2_ERROR := Y1 < 0 OR X1 < 0 OR Y2 < 0 OR X2 < 0 OR Y1 > 23 OR X1 > 79 OR Y2 > 23 OR X2 > 79;

END_FUNCTION

PROGRAM program0
	VAR
		X1 :	INT;
		Y1 :	INT;
		X2 :	INT;
		Y2 :	INT;
		CEIL5_OUT : BOOL;
	END_VAR

  	CEIL5_OUT := TN_SC_XY2_ERROR(X1, Y1, X2, Y2);
END_PROGRAM

CONFIGURATION Config0

  RESOURCE Res0 ON PLC
    TASK task0(INTERVAL := T#20ms,PRIORITY := 0);
    PROGRAM instance0 WITH task0 : program0;
  END_RESOURCE
END_CONFIGURATION

(* ---- 157-EVEN.ST ---- *)
FUNCTION BIT_OF_DWORD : BOOL
  VAR_INPUT
    IN : DWORD;
    N : INT;
  END_VAR

  BIT_OF_DWORD := (SHR(in,N) AND 16#00000001) > 0;
END_FUNCTION

FUNCTION EVEN:BOOL
	VAR_INPUT
		IN :	DINT;
	END_VAR

	even := NOT BIT_OF_DWORD(DINT_TO_DWORD(in),0);
END_FUNCTION

PROGRAM program0
  VAR
    LocalVar0 : DINT;
	  LocalOUT  : BOOL;
  END_VAR
  	LocalOUT := EVEN(LocalVar0);
END_PROGRAM

CONFIGURATION Config0
  RESOURCE Res0 ON PLC
    TASK task0(INTERVAL := T#20ms,PRIORITY := 0);
    PROGRAM instance0 WITH task0 : program0;
  END_RESOURCE
END_CONFIGURATION

(* ---- 159-BYTE_TO_TIME.ST ---- *)
FUNCTION _BYTE_TO_INT:INT
	VAR_INPUT
		IN :	BYTE;
	END_VAR

	_BYTE_TO_INT := USINT_TO_INT(BYTE_TO_USINT(IN));
END_FUNCTION

FUNCTION BYTE_TO_TIME2:TIME
	VAR_INPUT
		IN :	BYTE;
	END_VAR

	BYTE_TO_TIME2 := INT_TO_TIME(_BYTE_TO_INT(IN));
END_FUNCTION

PROGRAM program0
  VAR
    LocalVar0 : BYTE;
    CEIL5_OUT : TIME;
  END_VAR

  CEIL5_OUT := BYTE_TO_TIME2(LocalVar0);
END_PROGRAM

CONFIGURATION Config0

  RESOURCE Res0 ON PLC
    TASK task0(INTERVAL := T#20ms,PRIORITY := 0);
    PROGRAM instance0 WITH task0 : program0;
  END_RESOURCE
END_CONFIGURATION

(* ---- 16-DT_TO_DATE.ST ---- *)
FUNCTION _DT_TO_DATE_B:UDINT

	VAR_INPUT
		_INN :	UDINT;
	END_VAR

	_DT_TO_DATE_B := (_INN / UDINT#86400) * UDINT#86400;
END_FUNCTION

PROGRAM program0
	VAR
		_INN :	UDINT;
		OUT : UDINT;
	END_VAR

  OUT := _DT_TO_DATE_B(_INN);

END_PROGRAM

CONFIGURATION Config0
	RESOURCE Res0 ON PLC
		TASK task0(INTERVAL := T#20ms,PRIORITY := 0);
		PROGRAM instance0 WITH task0 : program0;
	END_RESOURCE
END_CONFIGURATION

(* ---- 161-TIMECHECK.ST ---- *)
FUNCTION TIMECHECK:BOOL

	VAR_INPUT
		TD :	UDINT;
		START :	UDINT;
		STOP :	UDINT;
	END_VAR

	IF stop < start THEN
		TIMECHECK := start <= TD OR  TD < stop;
	ELSE
		TIMECHECK := start <= TD AND TD < stop;
	END_IF;

END_FUNCTION

PROGRAM program0
  VAR
	TD :	UDINT;
	START :	UDINT;
	STOP :	UDINT;
    CEIL5_OUT : BOOL;
  END_VAR

  CEIL5_OUT := TIMECHECK(TD, START, STOP);
END_PROGRAM

CONFIGURATION Config0

  RESOURCE Res0 ON PLC
    TASK task0(INTERVAL := T#20ms,PRIORITY := 0);
    PROGRAM instance0 WITH task0 : program0;
  END_RESOURCE
END_CONFIGURATION

(* ---- 162-CIRCLE_SEG.ST ---- *)
FUNCTION CIRCLE_SEG:REAL
	VAR_INPUT
		RX :	REAL;
		HX :	REAL;
	END_VAR

	IF RX > 0.0 THEN
		CIRCLE_SEG := 2.0 * ACOS(1.0 - LIMIT(0.0, HX / RX, 2.0));
		CIRCLE_SEG := (CIRCLE_SEG - SIN(CIRCLE_SEG)) * RX * RX * 0.5;
	END_IF;
END_FUNCTION

PROGRAM program0
  VAR
    LocalVar0 : REAL;
	LocalVar1 : REAL;
	LocalOUT  : REAL;
  END_VAR
  	LocalOUT := CIRCLE_SEG(LocalVar0, LocalVar1);
END_PROGRAM

CONFIGURATION Config0
  RESOURCE Res0 ON PLC
    TASK task0(INTERVAL := T#20ms,PRIORITY := 0);
    PROGRAM instance0 WITH task0 : program0;
  END_RESOURCE
END_CONFIGURATION

(* ---- 163-GAUSS.ST ---- *)
FUNCTION GAUSS:REAL

	VAR_INPUT
		X :	REAL;
		U :	REAL;
		SI :	REAL;
	END_VAR

	VAR
		temp :	REAL;
		si_inv :	REAL;
	END_VAR

	temp := X - U;
	si_inv := 1.0  / si;
	GAUSS := EXP(Temp * Temp * si_inv * SI_inv * - 0.5) * 0.39894228 * si_inv;

END_FUNCTION

PROGRAM program0
  VAR
    X :	REAL;
	U :	REAL;
	SI :	REAL;
    LocalOUT  : REAL;
  END_VAR

  LocalOUT := GAUSS(X, U, SI);
END_PROGRAM

CONFIGURATION Config0
  RESOURCE Res0 ON PLC
    TASK task0(INTERVAL := T#20ms,PRIORITY := 0);
    PROGRAM instance0 WITH task0 : program0;
  END_RESOURCE
END_CONFIGURATION

(* ---- 164-BIT_LOAD_B.ST ---- *)
FUNCTION BIT_LOAD_B:BYTE
	VAR_INPUT
		IN :	BYTE;
		VAL :	BOOL;
		POS :	INT;
	END_VAR

	IF VAL THEN
		BIT_LOAD_B := in OR SHL(BYTE#1,pos);
	ELSE
		BIT_LOAD_B := in AND (NOT SHL(BYTE#1,pos));
	END_IF;
END_FUNCTION

PROGRAM program0
  VAR
    LocalVar0 : BYTE;
	LocalVar1 : BOOL;
	LocalVar2 : INT;
    LocalOUT  : BYTE;
  END_VAR

  LocalOUT := BIT_LOAD_B(LocalVar0, LocalVar1, LocalVar2);
END_PROGRAM

CONFIGURATION Config0
  RESOURCE Res0 ON PLC
    TASK task0(INTERVAL := T#20ms,PRIORITY := 0);
    PROGRAM instance0 WITH task0 : program0;
  END_RESOURCE
END_CONFIGURATION

(* ---- 165-BIT_LOAD_W.ST ---- *)
FUNCTION BIT_LOAD_W:WORD
	VAR_INPUT
		IN :	WORD;
		VAL :	BOOL;
		POS :	INT;
	END_VAR

	IF VAL THEN
		BIT_LOAD_W := in OR SHL(WORD#1,pos);
	ELSE
		BIT_LOAD_W := in AND (NOT SHL(WORD#1,pos));
	END_IF;
END_FUNCTION

PROGRAM program0
  VAR
    LocalVar0 : WORD;
	LocalVar1 : BOOL;
	LocalVar2 : INT;
    LocalOUT  : WORD;
  END_VAR

  LocalOUT := BIT_LOAD_W(LocalVar0, LocalVar1, LocalVar2);
END_PROGRAM

CONFIGURATION Config0
  RESOURCE Res0 ON PLC
    TASK task0(INTERVAL := T#20ms,PRIORITY := 0);
    PROGRAM instance0 WITH task0 : program0;
  END_RESOURCE
END_CONFIGURATION

(* ---- 166-MUX_4.ST ---- *)
FUNCTION MUX_4:BOOL

	VAR_INPUT
		D0 :	BOOL;
		D1 :	BOOL;
		D2 :	BOOL;
		D3 :	BOOL;
		A0 :	BOOL;
		A1 :	BOOL;
	END_VAR

	IF A1 THEN
		MUX_4 := SEL(A0, D2, D3);
	ELSE
		MUX_4 := SEL(A0, D0, D1);
	END_IF;

END_FUNCTION

PROGRAM program0
	VAR
		D0 :	BOOL;
		D1 :	BOOL;
		D2 :	BOOL;
		D3 :	BOOL;
		A0 :	BOOL;
		A1 :	BOOL;

		OUT : BOOL;
	END_VAR

	OUT := MUX_4(D0, D1, D2, D3, A0, A1);

END_PROGRAM

CONFIGURATION Config0

	RESOURCE Res0 ON PLC
		TASK task0(INTERVAL := T#20ms,PRIORITY := 0);
		PROGRAM instance0 WITH task0 : program0;
	END_RESOURCE

END_CONFIGURATION

(* ---- 167-BCDC_TO_INT.ST ---- *)
FUNCTION _BYTE_TO_INT:INT
	VAR_INPUT
		IN :	BYTE;
	END_VAR

	_BYTE_TO_INT := USINT_TO_INT(BYTE_TO_USINT(IN));

END_FUNCTION

FUNCTION BCDC_TO_INT:INT
	VAR_INPUT
		IN :	BYTE;
	END_VAR

	BCDC_TO_INT := _BYTE_TO_INT(in AND BYTE#16#0F) + (_BYTE_TO_INT(SHR(in,4)) * 10);
END_FUNCTION

PROGRAM program0
  VAR
    LocalVar0 : BYTE;
    LocalOUT  : INT;
  END_VAR

  LocalOUT := BCDC_TO_INT(LocalVar0);
END_PROGRAM

CONFIGURATION Config0
  RESOURCE Res0 ON PLC
    TASK task0(INTERVAL := T#20ms,PRIORITY := 0);
    PROGRAM instance0 WITH task0 : program0;
  END_RESOURCE
END_CONFIGURATION

(* ---- 168-BIT_COUNT.ST ---- *)
FUNCTION BIT_COUNT:INT

	VAR_INPUT
		IN :	DWORD;
	END_VAR

	VAR
		in_temp :	DWORD;
	END_VAR

	in_temp := IN;
	WHILE in_temp > DWORD#0 DO
		IF (in_temp AND DWORD#16#00000001) > DWORD#0 THEN Bit_Count := Bit_Count +1; END_IF;
		in_temp := SHR(in_temp,1);
	END_WHILE;

END_FUNCTION

PROGRAM program0
  VAR
    LocalVar0 : DWORD;
    LocalOUT  : INT;
  END_VAR

  LocalOUT := BIT_COUNT(LocalVar0);
END_PROGRAM

CONFIGURATION Config0
  RESOURCE Res0 ON PLC
    TASK task0(INTERVAL := T#20ms,PRIORITY := 0);
    PROGRAM instance0 WITH task0 : program0;
  END_RESOURCE
END_CONFIGURATION

(* ---- 169-LEAP_YEAR.ST ---- *)
FUNCTION LEAP_YEAR:BOOL

  VAR_INPUT
    YEAR :	INT;
  END_VAR

  IF (year MOD INT#400) = INT#00 THEN
    leap_year := TRUE;
  ELSIF (year MOD INT#100) = INT#00 THEN
    leap_year := FALSE;
  ELSIF (year MOD INT#04) = INT#00 THEN
    leap_year := TRUE;
  ELSE
    leap_year := FALSE;
  END_IF;

END_FUNCTION

PROGRAM program0
	VAR
		YEAR :	INT;
		OUT : BOOL;
	END_VAR

	OUT := LEAP_YEAR(YEAR);
END_PROGRAM

CONFIGURATION Config0

	RESOURCE Res0 ON PLC
		TASK task0(INTERVAL := T#20ms,PRIORITY := 0);
		PROGRAM instance0 WITH task0 : program0;
	END_RESOURCE

END_CONFIGURATION

(* ---- 17-INT_TO_TIME.ST ---- *)
FUNCTION _INT_TO_TIME:TIME

	VAR_INPUT
		IN :	INT;
	END_VAR

	_INT_TO_TIME := DINT_TO_TIME(INT_TO_DINT(IN));

END_FUNCTION

PROGRAM program0
	VAR
		IN :	INT;
		OUT : TIME;
	END_VAR

	OUT := _INT_TO_TIME(IN);
END_PROGRAM

CONFIGURATION Config0

	RESOURCE Res0 ON PLC
		TASK task0(INTERVAL := T#20ms,PRIORITY := 0);
		PROGRAM instance0 WITH task0 : program0;
	END_RESOURCE

END_CONFIGURATION

(* ---- 170-F_LIN2.ST ---- *)
FUNCTION F_LIN2:REAL
	VAR_INPUT
		X :	REAL;
		X1 :	REAL;
		Y1 :	REAL;
		X2 :	REAL;
		Y2 :	REAL;
	END_VAR

	F_LIN2 := (Y2 - Y1) / (X2 - X1) * (X - X1) + Y1;

END_FUNCTION

PROGRAM program0
  VAR
    LocalVar0 : REAL;
	LocalVar1 : REAL;
	LocalVar2 : REAL;
	LocalVar3 : REAL;
	LocalVar4 : REAL;
	  LocalOUT  : REAL;
  END_VAR
  	LocalOUT := F_LIN2(LocalVar0, LocalVar1, LocalVar2, LocalVar3, LocalVar4);
END_PROGRAM

CONFIGURATION Config0
  RESOURCE Res0 ON PLC
    TASK task0(INTERVAL := T#20ms,PRIORITY := 0);
    PROGRAM instance0 WITH task0 : program0;
  END_RESOURCE
END_CONFIGURATION

(* ---- 171-WORD_OF_DWORD.ST ---- *)
FUNCTION _BYTE_TO_INT:INT
	VAR_INPUT
		IN :	BYTE;
	END_VAR

	_BYTE_TO_INT := USINT_TO_INT(BYTE_TO_USINT(IN));
END_FUNCTION

FUNCTION WORD_OF_DWORD:WORD
	VAR_INPUT
		IN: DWORD;
		N :	BYTE;
	END_VAR
	WORD_OF_DWORD := DWORD_TO_WORD(SHR(in,_BYTE_TO_INT(SHL(n,4))));
END_FUNCTION

PROGRAM program0
  	VAR
		IN :	DWORD;
		N :	BYTE;
		CEIL5_OUT : WORD;
	  END_VAR

  	CEIL5_OUT := WORD_OF_DWORD(IN, N);
END_PROGRAM

CONFIGURATION Config0
  	RESOURCE Res0 ON PLC
    	TASK task0(INTERVAL := T#20ms,PRIORITY := 0);
    	PROGRAM instance0 WITH task0 : program0;
  	END_RESOURCE
END_CONFIGURATION

(* ---- 172-BIT_LOAD_DW.ST ---- *)
FUNCTION BIT_LOAD_DW:DWORD

	VAR_INPUT
		IN :	DWORD;
		VAL :	BOOL;
		POS :	INT;
	END_VAR

	IF val THEN
		BIT_LOAD_DW := in OR SHL(DWORD#1,pos);
	ELSE
		BIT_LOAD_DW := in AND (NOT SHL(DWORD#1,pos));
	END_IF;

END_FUNCTION

PROGRAM program0
  VAR
    LocalVar0 : DWORD;
	LocalVar1 : BOOL;
	LocalVar2 : INT;
    LocalOUT  : DWORD;
  END_VAR

  LocalOUT := BIT_LOAD_DW(LocalVar0, LocalVar1, LocalVar2);
END_PROGRAM

CONFIGURATION Config0
  RESOURCE Res0 ON PLC
    TASK task0(INTERVAL := T#20ms,PRIORITY := 0);
    PROGRAM instance0 WITH task0 : program0;
  END_RESOURCE
END_CONFIGURATION

(* ---- 173-DAYS_DELTA.ST ---- *)
FUNCTION DAYS_DELTA:DINT
	VAR_INPUT
		DATE_1 :	UDINT;
		DATE_2 :	UDINT;
	END_VAR
	IF DATE_1 > DATE_2 THEN
		DAYS_DELTA := - UDINT_TO_DINT((date_1 - date_2) / UDINT#86400);
	ELSE
		DAYS_DELTA :=   UDINT_TO_DINT((date_2 - date_1) / UDINT#86400);
	END_IF;
END_FUNCTION

PROGRAM program0
  VAR
    LocalVar0 : UDINT;
	LocalVar1 : UDINT;
	LocalOUT  : DINT;
  END_VAR
  	LocalOUT := DAYS_DELTA(LocalVar0, LocalVar1);
END_PROGRAM

CONFIGURATION Config0
  RESOURCE Res0 ON PLC
    TASK task0(INTERVAL := T#20ms,PRIORITY := 0);
    PROGRAM instance0 WITH task0 : program0;
  END_RESOURCE
END_CONFIGURATION

(* ---- 175-YEAR_BEGIN.ST ---- *)
FUNCTION _INT_TO_UDINT:UDINT
	VAR_INPUT
		IN :	INT;
	END_VAR

	_INT_TO_UDINT := DINT_TO_UDINT(INT_TO_DINT(IN));
END_FUNCTION

FUNCTION YEAR_BEGIN:UDINT
	VAR_INPUT
		Y :	INT;
	END_VAR
	year_begin := DWORD_TO_UDINT(SHR(UDINT_TO_DWORD(_INT_TO_UDINT(y) * UDINT#1461 - UDINT#2878169),2))*UDINT#86400;

END_FUNCTION

PROGRAM program0
  VAR
    Y : INT;
    CEIL5_OUT : UDINT;
  END_VAR

  CEIL5_OUT := YEAR_BEGIN(Y);
END_PROGRAM

CONFIGURATION Config0

  RESOURCE Res0 ON PLC
    TASK task0(INTERVAL := T#20ms,PRIORITY := 0);
    PROGRAM instance0 WITH task0 : program0;
  END_RESOURCE
END_CONFIGURATION

(* ---- 176-MUX_R4.ST ---- *)
FUNCTION MUX_R4:REAL

	VAR_INPUT
		IN0 :	REAL;
		IN1 :	REAL;
		IN2 :	REAL;
		IN3 :	REAL;
		A0 :	BOOL;
		A1 :	BOOL;
	END_VAR

	IF A1 THEN
		MUX_R4 := SEL(A0, IN2, IN3);
	ELSE
		MUX_R4 := SEL(A0, IN0, IN1);
	END_IF;

END_FUNCTION

PROGRAM program0
	VAR
		IN0 :	REAL;
		IN1 :	REAL;
		IN2 :	REAL;
		IN3 :	REAL;
		A0 :	BOOL;
		A1 :	BOOL;

		OUT : REAL;
	END_VAR

	OUT := MUX_R4(IN0, IN1, IN2, IN3, A0, A1);

END_PROGRAM

CONFIGURATION Config0

	RESOURCE Res0 ON PLC
		TASK task0(INTERVAL := T#20ms,PRIORITY := 0);
		PROGRAM instance0 WITH task0 : program0;
	END_RESOURCE

END_CONFIGURATION

(* ---- 177-RES_PT.ST ---- *)
FUNCTION RES_PT:REAL
	VAR_INPUT
		T :	REAL;
		R0 :	REAL;
	END_VAR

	VAR
		T2 :	REAL;
	END_VAR

	T2 := T * T;

	IF T >= 0.0 THEN
		RES_PT := R0 * ( 1.0 + 3.90802E-3 * T + -5.802E-7 * T2);
	ELSE
		RES_PT := R0 * ( 1.0 + 3.90802E-3 * T + -5.802E-7 * T2 + -4.27350E-12 * (T - 100.0) * T2 * T);
	END_IF;

END_FUNCTION

PROGRAM program0
  	VAR
		T :	REAL;
		R0 : REAL;
		CEIL5_OUT : REAL;
  	END_VAR

  	CEIL5_OUT := RES_PT(T, R0);
END_PROGRAM

CONFIGURATION Config0
	RESOURCE Res0 ON PLC
		TASK task0(INTERVAL := T#20ms,PRIORITY := 0);
		PROGRAM instance0 WITH task0 : program0;
	END_RESOURCE
END_CONFIGURATION

(* ---- 179-BYTE_OF_DWORD.ST ---- *)
FUNCTION _BYTE_TO_INT:INT
	VAR_INPUT
		IN :	BYTE;
	END_VAR

	_BYTE_TO_INT := USINT_TO_INT(BYTE_TO_USINT(IN));
END_FUNCTION

FUNCTION BYTE_OF_DWORD:BYTE
	VAR_INPUT
		IN :	DWORD;
		N :	BYTE;
	END_VAR
	BYTE_OF_DWORD := DWORD_TO_BYTE(SHR(in,_BYTE_TO_INT(SHL(n,3))));
END_FUNCTION

PROGRAM program0
  VAR
    LocalVar0 : DWORD;
	  LocalVar1 : BYTE;
    LocalOUT  : BYTE;
  END_VAR

  LocalOUT := BYTE_OF_DWORD(LocalVar0, LocalVar1);
END_PROGRAM

CONFIGURATION Config0
  RESOURCE Res0 ON PLC
    TASK task0(INTERVAL := T#20ms,PRIORITY := 0);
    PROGRAM instance0 WITH task0 : program0;
  END_RESOURCE
END_CONFIGURATION

(* ---- 185-SENSOR_INT.ST ---- *)
FUNCTION SENSOR_INT:REAL

	VAR_INPUT
		VOLTAGE :	REAL;
		CURRENT :	REAL;
		RP :	REAL;
		_RS :	REAL;
	END_VAR

	VAR
		RG :	REAL;
	END_VAR

	IF current <> 0.0 THEN
		RG := voltage / current;
		SENSOR_INT := RP * ( RG - _RS) / ( RP + _RS - RG);
	END_IF;

END_FUNCTION

PROGRAM program0

	VAR
		VOLTAGE :	REAL;
		CURRENT :	REAL;
		RP :	REAL;
		_RS :	REAL;
		CEIL5_OUT : REAL;
	END_VAR

	CEIL5_OUT := SENSOR_INT(VOLTAGE, CURRENT, RP, _RS);

END_PROGRAM

CONFIGURATION Config0

	RESOURCE Res0 ON PLC
		TASK task0(INTERVAL := T#20ms,PRIORITY := 0);
		PROGRAM instance0 WITH task0 : program0;
	END_RESOURCE

END_CONFIGURATION

(* ---- 186-DWORD_OF_BYTE.ST ---- *)
FUNCTION DWORD_OF_BYTE:DWORD
	VAR_INPUT
		B3 :	BYTE;
		B2 :	BYTE;
		B1 :	BYTE;
		B0 :	BYTE;
	END_VAR

	DWORD_OF_BYTE := SHL(SHL(SHL(BYTE_TO_DWORD(B3),8) OR BYTE_TO_DWORD(B2),8) OR BYTE_TO_DWORD(B1),8) OR BYTE_TO_DWORD(B0);

END_FUNCTION

PROGRAM program0
  VAR
    LocalVar0 : BYTE;
	LocalVar1 : BYTE;
	LocalVar2 : BYTE;
	LocalVar3 : BYTE;
	LocalOUT  : DWORD;
  END_VAR
  	LocalOUT := DWORD_OF_BYTE(LocalVar0, LocalVar1, LocalVar2, LocalVar3);
END_PROGRAM

CONFIGURATION Config0
  RESOURCE Res0 ON PLC
    TASK task0(INTERVAL := T#20ms,PRIORITY := 0);
    PROGRAM instance0 WITH task0 : program0;
  END_RESOURCE
END_CONFIGURATION

(* ---- 188-LANGEVIN.ST ---- *)
FUNCTION COTH:REAL

	VAR_INPUT
		X :	REAL;
	END_VAR

	IF X > 20.0 THEN
		COTH :=1.0;
	ELSIF X < -20.0 THEN
		COTH := -1.0;
	ELSE
		COTH := 1.0 + 2.0 / (EXP(X * 2.0) - 1.0);
	END_IF;

END_FUNCTION

FUNCTION LANGEVIN:REAL

	VAR_INPUT
		X :	REAL;
	END_VAR

	IF X = 0.0 THEN
		LANGEVIN := 0.0;
	ELSE
		LANGEVIN := COTH(X) - 1.0 / X;
	END_IF;

END_FUNCTION

PROGRAM program0
	VAR
		X :	REAL;
		OUT : REAL;
	END_VAR

	OUT := LANGEVIN(X);
END_PROGRAM

CONFIGURATION Config0

	RESOURCE Res0 ON PLC
		TASK task0(INTERVAL := T#20ms,PRIORITY := 0);
		PROGRAM instance0 WITH task0 : program0;
	END_RESOURCE

END_CONFIGURATION

(* ---- 19-ASINH.ST ---- *)
FUNCTION ASINH:REAL
	VAR_INPUT
		X :	REAL;
	END_VAR

	ASINH := LN(SQRT(X * X + 1.0)+X);
END_FUNCTION

PROGRAM program0
  VAR
    LocalVar0 : REAL;
    LocalOUT  : REAL;
  END_VAR

  LocalOUT := ASINH(LocalVar0);
END_PROGRAM

CONFIGURATION Config0
  RESOURCE Res0 ON PLC
    TASK task0(INTERVAL := T#20ms,PRIORITY := 0);
    PROGRAM instance0 WITH task0 : program0;
  END_RESOURCE
END_CONFIGURATION

(* ---- 192-D_TRUNC.ST ---- *)
FUNCTION D_TRUNC : DINT
  VAR_INPUT
    x : REAL;
  END_VAR

  D_TRUNC := REAL_TO_DINT(X);
  IF X > 0.0 THEN
  	IF DINT_TO_REAL(D_TRUNC) > X THEN D_TRUNC := D_TRUNC - DINT#1; END_IF;
  ELSE
  	IF DINT_TO_REAL(D_TRUNC) < X THEN D_TRUNC := D_TRUNC + DINT#1; END_IF;
  END_IF;
END_FUNCTION

PROGRAM program0
  VAR
    LocalVar0 : REAL;
    LocalVar1 : DINT;
    CEIL5_OUT : DINT;
  END_VAR

  CEIL5_OUT := D_TRUNC(LocalVar0);
  LocalVar1 := CEIL5_OUT;
END_PROGRAM

CONFIGURATION Config0

  RESOURCE Res0 ON PLC
    TASK task0(INTERVAL := T#20ms,PRIORITY := 0);
    PROGRAM instance0 WITH task0 : program0;
  END_RESOURCE
END_CONFIGURATION

(* ---- 193-SCALE_R.ST ---- *)
FUNCTION SCALE_R:REAL
	VAR_INPUT
		X :	REAL;
		I_LO :	REAL;
		I_HI :	REAL;
		O_LO :	REAL;
		O_HI :	REAL;
	END_VAR

	IF I_LO = I_HI THEN
		SCALE_R := O_LO;
	ELSE
		SCALE_R := (O_HI - O_LO) / (I_HI - I_LO) * (LIMIT(I_LO, X, I_HI) - I_LO) + O_LO;
	END_IF;

END_FUNCTION

PROGRAM program0

  	VAR
		X :	REAL;
		I_LO :	REAL;
		I_HI :	REAL;
		O_LO :	REAL;
		O_HI :	REAL;
		CEIL5_OUT : REAL;
  	END_VAR

  	CEIL5_OUT := SCALE_R(X, I_LO, I_HI, O_LO, O_HI);
END_PROGRAM

CONFIGURATION Config0

	RESOURCE Res0 ON PLC
		TASK task0(INTERVAL := T#20ms,PRIORITY := 0);
		PROGRAM instance0 WITH task0 : program0;
	END_RESOURCE

END_CONFIGURATION

(* ---- 194-BIT_LOAD_B2.ST ---- *)
FUNCTION BIT_LOAD_B2:BYTE
	VAR_INPUT
		I :	BYTE;
		D :	BOOL;
		P :	INT;
		N :	INT;
	END_VAR

	IF D THEN
		BIT_LOAD_B2 := ROL(SHR(BYTE#255, 8 - N) OR ROR(I, P), P);
	ELSE
		BIT_LOAD_B2 := ROL(SHL(BYTE#255, N) AND ROR(I, P), P);
	END_IF;
END_FUNCTION

PROGRAM program0
  VAR
    LocalVar0 : BYTE;
	LocalVar1 : BOOL;
	LocalVar2 : INT;
	LocalVar3 : INT;
    LocalOUT  : BYTE;
  END_VAR

  LocalOUT := BIT_LOAD_B2(LocalVar0, LocalVar1, LocalVar2, LocalVar3);
END_PROGRAM

CONFIGURATION Config0
  RESOURCE Res0 ON PLC
    TASK task0(INTERVAL := T#20ms,PRIORITY := 0);
    PROGRAM instance0 WITH task0 : program0;
  END_RESOURCE
END_CONFIGURATION

(* ---- 195-WORD_TO_RANGE.ST ---- *)
FUNCTION _WORD_TO_REAL:REAL
	VAR_INPUT
		IN :	WORD;
	END_VAR
	_WORD_TO_REAL := UINT_TO_REAL(WORD_TO_UINT(IN));
END_FUNCTION

FUNCTION WORD_TO_RANGE:REAL
	VAR_INPUT
		X :	WORD;
		LOW :	REAL;
		HIGH :	REAL;
	END_VAR
	WORD_TO_RANGE := (high - low) * _WORD_TO_REAL(X) * 0.00001525902189669640 + low;
END_FUNCTION

PROGRAM program0
  	VAR
		X :	WORD;
		LOW :	REAL;
		HIGH :	REAL;
		CEIL5_OUT : REAL;
	  END_VAR

  	CEIL5_OUT := WORD_TO_RANGE(X, LOW, HIGH);
END_PROGRAM

CONFIGURATION Config0
  	RESOURCE Res0 ON PLC
    	TASK task0(INTERVAL := T#20ms,PRIORITY := 0);
    	PROGRAM instance0 WITH task0 : program0;
  	END_RESOURCE
END_CONFIGURATION

(* ---- 196-BIT_LOAD_W2.ST ---- *)
FUNCTION BIT_LOAD_W2:WORD
	VAR_INPUT
		I :	WORD;
		D :	BOOL;
		P :	INT;
		N :	INT;
	END_VAR

	IF D THEN
		BIT_LOAD_W2 := ROL(SHR(WORD#16#FFFF, 16 - N) OR ROR(I, P), P);
	ELSE
		BIT_LOAD_W2 := ROL(SHL(WORD#16#FFFF, N) AND ROR(I, P), P);
	END_IF;
END_FUNCTION

PROGRAM program0
  VAR
    LocalVar0 : WORD;
	LocalVar1 : BOOL;
	LocalVar2 : INT;
	LocalVar3 : INT;
    LocalOUT  : WORD;
  END_VAR

  LocalOUT := BIT_LOAD_W2(LocalVar0, LocalVar1, LocalVar2, LocalVar3);
END_PROGRAM

CONFIGURATION Config0
  RESOURCE Res0 ON PLC
    TASK task0(INTERVAL := T#20ms,PRIORITY := 0);
    PROGRAM instance0 WITH task0 : program0;
  END_RESOURCE
END_CONFIGURATION

(* ---- 197-_REAL_TO_DWORD.ST ---- *)
FUNCTION _REAL_TO_DWORD: DWORD

  VAR_INPUT
    X :	REAL;
  END_VAR

  IF REAL_TO_DWORD(0.5) = DWORD#1 THEN
    _REAL_TO_DWORD := REAL_TO_DWORD(x);
  ELSIF X > 0.0 THEN
    _REAL_TO_DWORD := REAL_TO_DWORD(x+0.5);
  ELSIF X < 0.0 THEN
    _REAL_TO_DWORD := REAL_TO_DWORD(x-0.5);
  ELSE
    _REAL_TO_DWORD := DWORD#0;
  END_IF;
END_FUNCTION

PROGRAM program0
  VAR
    LocalVar0 : REAL;
    LocalOUT  : DWORD;
  END_VAR

  LocalOUT := _REAL_TO_DWORD(LocalVar0);
END_PROGRAM

CONFIGURATION Config0
  RESOURCE Res0 ON PLC
    TASK task0(INTERVAL := T#20ms,PRIORITY := 0);
    PROGRAM instance0 WITH task0 : program0;
  END_RESOURCE
END_CONFIGURATION

(* ---- 198-DAYS_IN_YEAR.ST ---- *)
FUNCTION LEAP_OF_DATE:BOOL

	VAR_INPUT
		IDATE :	UDINT;
	END_VAR

	LEAP_OF_DATE := SHL(UDINT_TO_DWORD((idate + UDINT#43200) / UDINT#31557600), 30) = DWORD#16#80000000;
END_FUNCTION

FUNCTION DAYS_IN_YEAR:INT
	VAR_INPUT
		IDATE :	UDINT;
	END_VAR

	IF LEAP_OF_DATE(IDATE) THEN
		DAYS_IN_YEAR := 366;
	ELSE
		DAYS_IN_YEAR := 365;
	END_IF;
END_FUNCTION

PROGRAM program0
  VAR
    LocalVar0 : UDINT;
	LocalOUT  : INT;
  END_VAR
  	LocalOUT := DAYS_IN_YEAR(LocalVar0);
END_PROGRAM

CONFIGURATION Config0
  RESOURCE Res0 ON PLC
    TASK task0(INTERVAL := T#20ms,PRIORITY := 0);
    PROGRAM instance0 WITH task0 : program0;
  END_RESOURCE
END_CONFIGURATION

(* ---- 20-SPHERE_V.ST ---- *)
FUNCTION SPHERE_V:REAL

	VAR_INPUT
		RX :	REAL;
	END_VAR

	sphere_V := 4.188790205 * Rx * RX * RX;

END_FUNCTION

PROGRAM program0

	VAR
		RX :	REAL;
		CEIL5_OUT : REAL;
	END_VAR

	CEIL5_OUT := SPHERE_V(RX);

END_PROGRAM

CONFIGURATION Config0

	RESOURCE Res0 ON PLC
		TASK task0(INTERVAL := T#20ms,PRIORITY := 0);
		PROGRAM instance0 WITH task0 : program0;
	END_RESOURCE

END_CONFIGURATION

(* ---- 200-_REAL_TO_DINT.ST ---- *)
FUNCTION _REAL_TO_DINT:DINT
  VAR_INPUT
    X :	REAL;
  END_VAR

  IF REAL_TO_DINT(0.5) = DINT#1 THEN
    _REAL_TO_DINT := REAL_TO_DINT(x);
    RETURN;
  END_IF;

  IF X > 0.0 THEN
    _REAL_TO_DINT := REAL_TO_DINT(x+0.5);
  ELSIF X < 0.0 THEN
    _REAL_TO_DINT := REAL_TO_DINT(x-0.5);
  ELSE
    _REAL_TO_DINT := DINT#0;
  END_IF;
END_FUNCTION

PROGRAM program0
  VAR
    LocalVar0 : REAL;
	  LocalOUT  : DINT;
  END_VAR

  LocalOUT := _REAL_TO_DINT(LocalVar0);
END_PROGRAM

CONFIGURATION Config0
  RESOURCE Res0 ON PLC
    TASK task0(INTERVAL := T#20ms,PRIORITY := 0);
    PROGRAM instance0 WITH task0 : program0;
  END_RESOURCE
END_CONFIGURATION

(* ---- 203-RANGE_TO_BYTE.ST ---- *)
FUNCTION TRUNC_REAL:REAL

	VAR_INPUT
		IN :	REAL;
	END_VAR

	TRUNC_REAL := UDINT_TO_REAL(DINT_TO_UDINT(TRUNC(IN)));
END_FUNCTION

FUNCTION RANGE_TO_BYTE:BYTE

	VAR_INPUT
		X :	REAL;
		LOW :	REAL;
		HIGH :	REAL;
	END_VAR

	Range_to_Byte := REAL_TO_BYTE(TRUNC_REAL((LIMIT(low,X,high)-low) * 255.0 / (high - low)));

END_FUNCTION

PROGRAM program0

	VAR
		X :	REAL;
		LOW :	REAL;
		HIGH :	REAL;

        OUT :	BYTE;
	END_VAR
	OUT := RANGE_TO_BYTE(X, LOW, HIGH);

END_PROGRAM

CONFIGURATION Config0

	RESOURCE Res0 ON PLC
		TASK task0(INTERVAL := T#20ms,PRIORITY := 0);
		PROGRAM instance0 WITH task0 : program0;
	END_RESOURCE

END_CONFIGURATION

(* ---- 204-RANGE_TO_WORD.ST ---- *)
FUNCTION TRUNC_REAL:REAL

	VAR_INPUT
		IN :	REAL;
	END_VAR

	TRUNC_REAL := UDINT_TO_REAL(DINT_TO_UDINT(TRUNC(IN)));
END_FUNCTION

FUNCTION RANGE_TO_WORD:WORD

	VAR_INPUT
		X :	REAL;
		LOW :	REAL;
		HIGH :	REAL;
	END_VAR

	Range_to_Word := REAL_TO_WORD(TRUNC_REAL((LIMIT(low,X,high)-low) * 65535.0 / (high - low)));

END_FUNCTION

PROGRAM program0

	VAR
		X :	REAL;
		LOW :	REAL;
		HIGH :	REAL;

        OUT :	WORD;
	END_VAR
	OUT := RANGE_TO_WORD(X, LOW, HIGH);

END_PROGRAM

CONFIGURATION Config0

	RESOURCE Res0 ON PLC
		TASK task0(INTERVAL := T#20ms,PRIORITY := 0);
		PROGRAM instance0 WITH task0 : program0;
	END_RESOURCE

END_CONFIGURATION

(* ---- 205-REFLECT.ST ---- *)
FUNCTION REFLECT:DWORD
	VAR_INPUT
		D :	DWORD;
		L :	INT;
	END_VAR

	VAR
		i :	INT;
		_d :	DWORD;
	END_VAR

	REFLECT := DWORD#0;
	_d := D;
	FOR i := 1 TO L DO
		REFLECT := SHL(REFLECT, 1) OR BOOL_TO_DWORD((_d AND DWORD#2#0000_0001) > DWORD#0); (* D.0 *)
		_d := SHR(_d, 1);
	END_FOR;
	REFLECT := REFLECT OR SHL(_d, L);
END_FUNCTION

PROGRAM program0
  VAR
    LocalVar0 : DWORD;
	LocalVar1 : INT;
	LocalOUT  : DWORD;
  END_VAR
  	LocalOUT := REFLECT(LocalVar0, LocalVar1);
END_PROGRAM

CONFIGURATION Config0
  RESOURCE Res0 ON PLC
    TASK task0(INTERVAL := T#20ms,PRIORITY := 0);
    PROGRAM instance0 WITH task0 : program0;
  END_RESOURCE
END_CONFIGURATION

(* ---- 206-_REAL_TO_UDINT.ST ---- *)
FUNCTION _REAL_TO_UDINT:UDINT
  VAR_INPUT
    X :	REAL;
  END_VAR

  IF REAL_TO_UDINT(0.5) = UDINT#1 THEN
    _REAL_TO_UDINT := REAL_TO_UDINT(x);
  ELSIF X > 0.0 THEN
    _REAL_TO_UDINT := REAL_TO_UDINT(x+0.5);
  ELSIF X < 0.0 THEN
    _REAL_TO_UDINT := REAL_TO_UDINT(x-0.5);
  ELSE
    _REAL_TO_UDINT := UDINT#0;
  END_IF;
END_FUNCTION

PROGRAM program0
    VAR
      LocalVar0 : REAL;
      LocalOUT  : UDINT;
    END_VAR

    LocalOUT := _REAL_TO_UDINT(LocalVar0);
END_PROGRAM

CONFIGURATION Config0
    RESOURCE Res0 ON PLC
      TASK task0(INTERVAL := T#20ms,PRIORITY := 0);
      PROGRAM instance0 WITH task0 : program0;
    END_RESOURCE
END_CONFIGURATION

(* ---- 208-BETA.ST ---- *)
FUNCTION GAMMA:REAL
	VAR_INPUT
		X :	REAL;
	END_VAR

	IF x > 0.0 THEN
		GAMMA := SQRT(6.28318530717958647692528676655900576 / X) * EXPT(0.367879441171442 * (x + 1.0 / (12.0 * x - 0.1 / X)), X);
	END_IF;
END_FUNCTION

FUNCTION BETA:REAL

	VAR_INPUT
		X :	REAL;
		Y :	REAL;
	END_VAR

	BETA := GAMMA(X)*GAMMA(Y) / GAMMA(x+y);

END_FUNCTION

PROGRAM program0
  VAR
    LocalVar0 : REAL;
	LocalVar1 : REAL;
    LocalOUT  : REAL;
  END_VAR

  LocalOUT := BETA(LocalVar0, LocalVar1);
END_PROGRAM

CONFIGURATION Config0
  RESOURCE Res0 ON PLC
    TASK task0(INTERVAL := T#20ms,PRIORITY := 0);
    PROGRAM instance0 WITH task0 : program0;
  END_RESOURCE
END_CONFIGURATION

(* ---- 209-ISC_LOWER.ST ---- *)
FUNCTION SETUP_EXTENDED_ASCII:BOOL

	VAR_INPUT
		X :	BOOL;
	END_VAR

	SETUP_EXTENDED_ASCII := X OR TRUE;

END_FUNCTION

FUNCTION ISC_LOWER:BOOL

	VAR_INPUT
		IN :	BYTE;
	END_VAR

	IF SETUP_EXTENDED_ASCII(FALSE) THEN
		ISC_LOWER := ((in > BYTE#96) AND (in < BYTE#123)) OR ((in > BYTE#222) AND (in <> BYTE#247));
	ELSE
		ISC_LOWER := ((in > BYTE#96) AND (in < BYTE#123));
	END_IF;

END_FUNCTION

PROGRAM program0
	VAR
		IN : BYTE;
		OUT : BOOL;
	END_VAR

	OUT := ISC_LOWER(IN);
END_PROGRAM

CONFIGURATION Config0

	RESOURCE Res0 ON PLC
		TASK task0(INTERVAL := T#20ms,PRIORITY := 0);
		PROGRAM instance0 WITH task0 : program0;
	END_RESOURCE

END_CONFIGURATION

(* ---- 21-AGDF.ST ---- *)
FUNCTION AGDF:REAL
	VAR_INPUT
		X :	REAL;
	END_VAR

	AGDF := LN((1.0 + SIN(X)) / COS(X));
END_FUNCTION

PROGRAM program0
  VAR
    LocalVar0 : REAL;
    LocalOUT  : REAL;
  END_VAR

  LocalOUT := AGDF(LocalVar0);
END_PROGRAM

CONFIGURATION Config0
  RESOURCE Res0 ON PLC
    TASK task0(INTERVAL := T#20ms,PRIORITY := 0);
    PROGRAM instance0 WITH task0 : program0;
  END_RESOURCE
END_CONFIGURATION

(* ---- 210-BIT_LOAD_DW2.ST ---- *)
FUNCTION BIT_LOAD_DW2:DWORD
	VAR_INPUT
		I :	DWORD;
		D :	BOOL;
		P :	INT;
		N :	INT;
	END_VAR

	IF D THEN
		BIT_LOAD_DW2 := ROL(SHR(DWORD#16#FFFFFFFF, 32 - N) OR ROR(I, P), P);
	ELSE
		BIT_LOAD_DW2 := ROL(SHL(DWORD#16#FFFFFFFF, N) AND ROR(I, P), P);
	END_IF;

END_FUNCTION

PROGRAM program0
  VAR
    LocalVar0 : DWORD;
	LocalVar1 : BOOL;
	LocalVar2 : INT;
	LocalVar3 : INT;
    LocalOUT  : DWORD;
  END_VAR

  LocalOUT := BIT_LOAD_DW2(LocalVar0, LocalVar1, LocalVar2, LocalVar3);
END_PROGRAM

CONFIGURATION Config0
  RESOURCE Res0 ON PLC
    TASK task0(INTERVAL := T#20ms,PRIORITY := 0);
    PROGRAM instance0 WITH task0 : program0;
  END_RESOURCE
END_CONFIGURATION

(* ---- 212-MID3.ST ---- *)
FUNCTION MID3:REAL

	VAR_INPUT
		IN1 :	REAL;
		IN2 :	REAL;
		IN3 :	REAL;
	END_VAR

	VAR
		_IN1 :	REAL;
		_IN2 :	REAL;
		_IN3 :	REAL;
	END_VAR

	_IN1 := IN1;
	_IN2 := IN2;
	_IN3 := IN3;

	IF _IN1 > _IN2 THEN MID3 := _IN1; _IN1 := _IN2; _IN2 := MID3; END_IF;
	IF _IN2 > _IN3 THEN _IN2 := _IN3; END_IF;
	MID3 := SEL(_IN1 > _IN2, _IN2, _IN1);

END_FUNCTION

PROGRAM program0
	VAR
		IN1 :	REAL;
		IN2 :	REAL;
		IN3 :	REAL;

		OUT : REAL;
	END_VAR

	OUT := MID3(IN1, IN2, IN3);

END_PROGRAM

CONFIGURATION Config0

	RESOURCE Res0 ON PLC
		TASK task0(INTERVAL := T#20ms,PRIORITY := 0);
		PROGRAM instance0 WITH task0 : program0;
	END_RESOURCE

END_CONFIGURATION

(* ---- 213-BYTE_TO_RANGE.ST ---- *)
FUNCTION _BYTE_TO_REAL:REAL
	VAR_INPUT
		IN :	BYTE;
	END_VAR

	_BYTE_TO_REAL := USINT_TO_REAL(BYTE_TO_USINT(IN));
END_FUNCTION

FUNCTION BYTE_TO_RANGE:REAL
	VAR_INPUT
		X :	BYTE;
		LOW :	REAL;
		HIGH :	REAL;
	END_VAR

	Byte_to_Range := (high - low) * _BYTE_TO_REAL(X) / 255.0 + low;
END_FUNCTION

PROGRAM program0
  VAR
    LocalVar0 : BYTE;
    LocalVar1 : REAL;
	LocalVar2 : REAL;
    CEIL5_OUT : REAL;
  END_VAR

  CEIL5_OUT := BYTE_TO_RANGE(LocalVar0, LocalVar1, LocalVar2);
END_PROGRAM

CONFIGURATION Config0

  RESOURCE Res0 ON PLC
    TASK task0(INTERVAL := T#20ms,PRIORITY := 0);
    PROGRAM instance0 WITH task0 : program0;
  END_RESOURCE
END_CONFIGURATION

(* ---- 216-MODR.ST ---- *)
FUNCTION FLOOR2 : DINT
	VAR_INPUT
		x : REAL;
	END_VAR

	FLOOR2 := REAL_TO_DINT(X);
	IF DINT_TO_REAL(FLOOR2) > X THEN
		FLOOR2 := FLOOR2 - DINT#1;
	END_IF;

END_FUNCTION

FUNCTION MODR: REAL

	VAR_INPUT
		IN :	REAL;
		DIVI :	REAL;
	END_VAR

	IF divi = 0.0 THEN
		MODR := 0.0;
	ELSE
		MODR := in - DINT_TO_REAL(FLOOR2(in / divi)) * divi;
	END_IF;

END_FUNCTION

PROGRAM program0

  	VAR
		IN :	REAL;
		DIVI :	REAL;
		CEIL5_OUT : REAL;
  	END_VAR

  	CEIL5_OUT := MODR(IN, DIVI);
END_PROGRAM

CONFIGURATION Config0

  RESOURCE Res0 ON PLC
    TASK task0(INTERVAL := T#20ms,PRIORITY := 0);
    PROGRAM instance0 WITH task0 : program0;
  END_RESOURCE
END_CONFIGURATION

(* ---- 218-CTRL_IN.ST ---- *)
FUNCTION DEAD_ZONE:REAL

	VAR_INPUT
		X :	REAL;
		L :	REAL;
	END_VAR

	IF ABS(x) > L THEN
		dead_zone := X;
	ELSE
		DEAD_ZONE := 0.0;
	END_IF;

END_FUNCTION

FUNCTION CTRL_IN:REAL
	VAR_INPUT
		SET_POINT :	REAL;
		ACTUAL :	REAL;
		NOISE :	REAL;
	END_VAR
	CTRL_IN := DEAD_ZONE(SET_POINT - ACTUAL, NOISE);
END_FUNCTION

PROGRAM program0
  VAR
    LocalVar0 : REAL;
	LocalVar1 : REAL;
	LocalVar2 : REAL;
	LocalOUT  : REAL;
  END_VAR
  	LocalOUT := CTRL_IN(LocalVar0, LocalVar1, LocalVar2);
END_PROGRAM

CONFIGURATION Config0
  RESOURCE Res0 ON PLC
    TASK task0(INTERVAL := T#20ms,PRIORITY := 0);
    PROGRAM instance0 WITH task0 : program0;
  END_RESOURCE
END_CONFIGURATION

(* ---- 22-HOUR.ST ---- *)
FUNCTION HOUR:INT
	VAR_INPUT
		ITOD :	UDINT;
	END_VAR
	hour := UDINT_TO_INT(itod / UDINT#3600000);
END_FUNCTION

PROGRAM program0
  VAR
	  ITOD :	UDINT;
    CEIL5_OUT : INT;
  END_VAR

  CEIL5_OUT := HOUR(ITOD);
END_PROGRAM

CONFIGURATION Config0

  RESOURCE Res0 ON PLC
    TASK task0(INTERVAL := T#20ms,PRIORITY := 0);
    PROGRAM instance0 WITH task0 : program0;
  END_RESOURCE
END_CONFIGURATION

(* ---- 221-ISC_UPPER.ST ---- *)
FUNCTION SETUP_EXTENDED_ASCII:BOOL

	VAR_INPUT
		X :	BOOL;
	END_VAR

	SETUP_EXTENDED_ASCII := X OR TRUE;

END_FUNCTION

FUNCTION ISC_UPPER:BOOL

	VAR_INPUT
		IN :	BYTE;
	END_VAR

	IF SETUP_EXTENDED_ASCII(FALSE) THEN
		ISC_UPPER :=  ((in > BYTE#64) AND (in < BYTE#91)) OR (((in > BYTE#191) AND (in < BYTE#223)) AND (in <> BYTE#215));
	ELSE
		ISC_UPPER := ((in > BYTE#64) AND (in < BYTE#91));
	END_IF;

END_FUNCTION

PROGRAM program0
	VAR
		IN : BYTE;
		OUT : BOOL;
	END_VAR

	OUT := ISC_UPPER(IN);
END_PROGRAM

CONFIGURATION Config0

	RESOURCE Res0 ON PLC
		TASK task0(INTERVAL := T#20ms,PRIORITY := 0);
		PROGRAM instance0 WITH task0 : program0;
	END_RESOURCE

END_CONFIGURATION

(* ---- 224-_ARRAY_ABS.ST ---- *)
TYPE
	oscat_pt_ARRAY: ARRAY [1..100] OF REAL;
END_TYPE

FUNCTION _ARRAY_ABS : BOOL
	VAR_IN_OUT
		PT : oscat_pt_ARRAY;
	END_VAR

	VAR_INPUT
		SIZE :	UINT;
	END_VAR

	VAR
		i :	INT;
		stop :	INT;
	END_VAR

	stop := LIMIT_INT(1,UINT_TO_INT(size),1000);
	FOR i := 1 TO stop DO
		pt[i] := ABS(pt[i]);
	END_FOR;

	_ARRAY_ABS := TRUE;

END_FUNCTION

PROGRAM program0
  VAR
    LocalVar0 : oscat_pt_ARRAY;
    LocalVar1 : UINT;
	LocalOUT  : BOOL;
  END_VAR

  LocalOUT := _ARRAY_ABS(LocalVar0, LocalVar1);
END_PROGRAM

CONFIGURATION Config0
  RESOURCE Res0 ON PLC
    TASK task0(INTERVAL := T#20ms,PRIORITY := 0);
    PROGRAM instance0 WITH task0 : program0;
  END_RESOURCE
END_CONFIGURATION

(* ---- 226-TANK_VOL1.ST ---- *)
FUNCTION CIRCLE_SEG:REAL
	VAR_INPUT
		RX :	REAL;
		HX :	REAL;
	END_VAR

	IF RX > 0.0 THEN
		CIRCLE_SEG := 2.0 * ACOS(1.0 - LIMIT(0.0, HX / RX, 2.0));
		CIRCLE_SEG := (CIRCLE_SEG - SIN(CIRCLE_SEG)) * RX * RX * 0.5;
	END_IF;
END_FUNCTION

FUNCTION TANK_VOL1:REAL

	VAR_INPUT
		TR :	REAL;
		TL :	REAL;
		H :	REAL;
	END_VAR

	TANK_VOL1 := CIRCLE_SEG(TR, H) * TL;

END_FUNCTION

PROGRAM program0
  VAR
    TR :	REAL;
	TL :	REAL;
	H :	REAL;
    CEIL5_OUT : REAL;
  END_VAR

  CEIL5_OUT := TANK_VOL1(TR, TL, H);
END_PROGRAM

CONFIGURATION Config0

  RESOURCE Res0 ON PLC
    TASK task0(INTERVAL := T#20ms,PRIORITY := 0);
    PROGRAM instance0 WITH task0 : program0;
  END_RESOURCE
END_CONFIGURATION

(* ---- 229-ERF.ST ---- *)
FUNCTION SGN : INT
  VAR_INPUT
    x : REAL;
  END_VAR

  IF X > 0.0 THEN
  	sgn := 1;
  ELSIF X < 0.0 THEN
  	sgn := -1;
  ELSE
  	sgn := 0;
  END_IF;
END_FUNCTION

FUNCTION ERF:REAL

	VAR_INPUT
		X :	REAL;
	END_VAR

	VAR
		x2 :	REAL;
		ax2 :	REAL;
	END_VAR

	x2 := X*X;
	ax2 := 0.147 * x2 + 1.0;
	ERF := SQRT(1.0 - EXP(-X2 * ((0.27323954473516 + aX2)/(ax2)))) * INT_TO_REAL(SGN(x));

END_FUNCTION

PROGRAM program0
  VAR
    LocalVar0 : REAL;
	  LocalOUT  : REAL;
  END_VAR
  	LocalOUT := ERF(LocalVar0);
END_PROGRAM

CONFIGURATION Config0
  RESOURCE Res0 ON PLC
    TASK task0(INTERVAL := T#20ms,PRIORITY := 0);
    PROGRAM instance0 WITH task0 : program0;
  END_RESOURCE
END_CONFIGURATION

(* ---- 23-ACOSH.ST ---- *)
FUNCTION ACOSH:REAL
	VAR_INPUT
		X :	REAL;
	END_VAR
	ACOSH := LN(SQRT(X * X - 1.0) + X);

END_FUNCTION

PROGRAM program0
  VAR
    LocalVar0 : REAL;
    LocalOUT  : REAL;
  END_VAR

  LocalOUT := ACOSH(LocalVar0);
END_PROGRAM

CONFIGURATION Config0
  RESOURCE Res0 ON PLC
    TASK task0(INTERVAL := T#20ms,PRIORITY := 0);
    PROGRAM instance0 WITH task0 : program0;
  END_RESOURCE
END_CONFIGURATION

(* ---- 230-DAY_OF_YEAR.ST ---- *)
FUNCTION DAY_OF_YEAR:INT
	VAR_INPUT
		IDATE :	DATE;
	END_VAR

	DAY_OF_YEAR := UDINT_TO_INT((DATE_TO_UDINT(idate) / UDINT#86400) MOD UDINT#1461);
	IF DAY_OF_YEAR > 729 THEN
		IF DAY_OF_YEAR > 1095 THEN DAY_OF_YEAR := DAY_OF_YEAR - 1095; ELSE DAY_OF_YEAR := DAY_OF_YEAR - 729; END_IF;
	ELSIF DAY_OF_YEAR > 364 THEN
		DAY_OF_YEAR := DAY_OF_YEAR - 364;
	ELSE
		DAY_OF_YEAR := DAY_OF_YEAR + 1;
	END_IF;
END_FUNCTION

PROGRAM program0
  VAR
    LocalVar0 : DATE;
	LocalOUT  : INT;
  END_VAR
  	LocalOUT := DAY_OF_YEAR(LocalVar0);
END_PROGRAM

CONFIGURATION Config0
  RESOURCE Res0 ON PLC
    TASK task0(INTERVAL := T#20ms,PRIORITY := 0);
    PROGRAM instance0 WITH task0 : program0;
  END_RESOURCE
END_CONFIGURATION

(* ---- 231-PARITY.ST ---- *)
FUNCTION BIT_OF_DWORD : BOOL

	VAR_INPUT
		IN : DWORD;
		N : INT;
	END_VAR

	BIT_OF_DWORD := (SHR(in,N) AND 16#00000001) > 0;

END_FUNCTION

FUNCTION PARITY:BOOL

	VAR_INPUT
		IN :	DWORD;
	END_VAR

	VAR
		in2 :	DWORD;
	END_VAR

	in2:=in;
	WHILE in2 > DWORD#0 DO
		parity := parity XOR BIT_OF_DWORD(in2,0) XOR BIT_OF_DWORD(in2,1) XOR BIT_OF_DWORD(in2,2) XOR BIT_OF_DWORD(in2,3);
		in2 := SHR(in2,4);
	END_WHILE;

END_FUNCTION

PROGRAM program0
	VAR
		IN : DWORD;
		OUT : BOOL;
	END_VAR

	OUT := PARITY(IN);
END_PROGRAM

CONFIGURATION Config0

	RESOURCE Res0 ON PLC
		TASK task0(INTERVAL := T#20ms,PRIORITY := 0);
		PROGRAM instance0 WITH task0 : program0;
	END_RESOURCE

END_CONFIGURATION

(* ---- 234-DEW_TEMP.ST ---- *)
FUNCTION EXP10 : REAL
  VAR_INPUT
    x : REAL;
  END_VAR

  exp10 := EXP(X * 2.30258509299405);
  (* from OSCAT library; www.oscat.de  *)
END_FUNCTION

FUNCTION DEW_TEMP:REAL

VAR_INPUT
	RH :	REAL;
	T :	REAL;
END_VAR

	VAR
		V :	REAL;
	END_VAR

	IF rh > 0.0 THEN

		V := LOG(RH * 0.01 * EXP10((7.5*T) / (237.3+T)));
		DEW_TEMP := 237.3*V / (7.5-V);
	ELSE
		DEW_TEMP:= -273.15;
	END_IF;

END_FUNCTION

PROGRAM program0
	VAR
		RH :	REAL;
		T :	REAL;
		CEIL5_OUT : REAL;
	END_VAR

  	CEIL5_OUT := DEW_TEMP(RH, T);
END_PROGRAM

CONFIGURATION Config0

  RESOURCE Res0 ON PLC
    TASK task0(INTERVAL := T#20ms,PRIORITY := 0);
    PROGRAM instance0 WITH task0 : program0;
  END_RESOURCE
END_CONFIGURATION

(* ---- 237-TO_UPPER.ST ---- *)
FUNCTION SETUP_EXTENDED_ASCII:BOOL
	VAR_INPUT
		X :	BOOL;
	END_VAR

	SETUP_EXTENDED_ASCII := X OR TRUE;
END_FUNCTION

FUNCTION TO_UPPER:BYTE

	VAR_INPUT
		IN :	BYTE;
	END_VAR

	IF in > BYTE#96 AND in < BYTE#123 THEN
	TO_UPPER := in AND BYTE#16#DF;
	ELSIF in > BYTE#223 AND in <> BYTE#247 AND in <> BYTE#255 AND SETUP_EXTENDED_ASCII(FALSE) THEN
	TO_UPPER := in AND BYTE#16#DF;
	ELSE
	TO_UPPER := in;
	END_IF;

END_FUNCTION

PROGRAM program0
  VAR
	IN :	BYTE;
    CEIL5_OUT : BYTE;
  END_VAR

  CEIL5_OUT := TO_UPPER(IN);
END_PROGRAM

CONFIGURATION Config0

  RESOURCE Res0 ON PLC
    TASK task0(INTERVAL := T#20ms,PRIORITY := 0);
    PROGRAM instance0 WITH task0 : program0;
  END_RESOURCE
END_CONFIGURATION

(* ---- 239-TO_LOWER.ST ---- *)
FUNCTION SETUP_EXTENDED_ASCII:BOOL

	VAR_INPUT
		X :	BOOL;
	END_VAR

	SETUP_EXTENDED_ASCII := X OR TRUE;
END_FUNCTION

FUNCTION TO_LOWER:BYTE

	VAR_INPUT
		IN :	BYTE;
	END_VAR

	IF in > BYTE#64 AND in < BYTE#91 THEN
	TO_LOWER := in OR BYTE#16#20;
	ELSIF (in > BYTE#191 AND in < BYTE#223) AND in <> BYTE#215 AND SETUP_EXTENDED_ASCII(FALSE) THEN
	TO_LOWER := in OR BYTE#16#20;
	ELSE
	TO_LOWER := in;
	END_IF;

END_FUNCTION

PROGRAM program0
  VAR
	IN :	BYTE;
    CEIL5_OUT : BYTE;
  END_VAR

  CEIL5_OUT := TO_LOWER(IN);
END_PROGRAM

CONFIGURATION Config0

  RESOURCE Res0 ON PLC
    TASK task0(INTERVAL := T#20ms,PRIORITY := 0);
    PROGRAM instance0 WITH task0 : program0;
  END_RESOURCE
END_CONFIGURATION

(* ---- 24-TOD_TO_REAL.ST ---- *)
FUNCTION TOD_TO_REAL2:REAL
	VAR_INPUT
		IN :	UDINT;
	END_VAR
	TOD_TO_REAL2 := UDINT_TO_REAL(IN);
END_FUNCTION

PROGRAM program0
  VAR
	IN :	UDINT;
    CEIL5_OUT : REAL;
  END_VAR

  CEIL5_OUT := TOD_TO_REAL2(IN);
END_PROGRAM

CONFIGURATION Config0

  RESOURCE Res0 ON PLC
    TASK task0(INTERVAL := T#20ms,PRIORITY := 0);
    PROGRAM instance0 WITH task0 : program0;
  END_RESOURCE
END_CONFIGURATION

(* ---- 242-FACT.ST ---- *)
FUNCTION FACT:DINT

	VAR_INPUT
		X :	INT;
	END_VAR

	CASE X OF
	00: FACT := DINT#1;
	01: FACT := DINT#1;
	02: FACT := DINT#2;
	03: FACT := DINT#6;
	04: FACT := DINT#24;
	05: FACT := DINT#120;
	06: FACT := DINT#720;
	07: FACT := DINT#5040;
	08: FACT := DINT#40320;
	09: FACT := DINT#362880;
	10: FACT := DINT#3628800;
	11: FACT := DINT#39916800;
	12: FACT := DINT#479001600;
	ELSE
		FACT := DINT#-1;
	END_CASE;

END_FUNCTION

PROGRAM program0
  VAR
    LocalVar0 : INT;
	LocalOUT  : DINT;
  END_VAR
  	LocalOUT := FACT(LocalVar0);
END_PROGRAM

CONFIGURATION Config0
  RESOURCE Res0 ON PLC
    TASK task0(INTERVAL := T#20ms,PRIORITY := 0);
    PROGRAM instance0 WITH task0 : program0;
  END_RESOURCE
END_CONFIGURATION

(* ---- 246-_ARRAY_ADD.ST ---- *)
TYPE
	oscat_pt_ARRAY: ARRAY [1..100] OF REAL;
END_TYPE

FUNCTION _ARRAY_ADD:	BOOL
	VAR_IN_OUT
		PT :	oscat_pt_ARRAY;
	END_VAR
	VAR_INPUT
		SIZE :	UINT;
		X :	REAL;
	END_VAR
	VAR
		i :	INT;
		stop :	INT;
	END_VAR

	stop :=LIMIT_INT(1,UINT_TO_INT(size),1000);
	FOR i := 1 TO stop DO
		pt[i] := pt[i] + X;
	END_FOR;
	_ARRAY_ADD := TRUE;

END_FUNCTION

PROGRAM program0
  VAR
    LocalVar0 : oscat_pt_ARRAY;
    LocalVar1 : UINT;
	LocalVar2 : REAL;
	LocalOUT  : BOOL;
  END_VAR

  LocalOUT := _ARRAY_ADD(LocalVar0, LocalVar1, LocalVar2);
END_PROGRAM

CONFIGURATION Config0
  RESOURCE Res0 ON PLC
    TASK task0(INTERVAL := T#20ms,PRIORITY := 0);
    PROGRAM instance0 WITH task0 : program0;
  END_RESOURCE
END_CONFIGURATION

(* ---- 248-LTIME_TO_UTC.ST ---- *)
FUNCTION _INT_TO_UDINT:UDINT
	VAR_INPUT
		IN :	INT;
	END_VAR

	_INT_TO_UDINT := DINT_TO_UDINT(INT_TO_DINT(IN));
END_FUNCTION

FUNCTION LTIME_TO_UTC:UDINT

	VAR_INPUT
		LTIME :	UDINT;
		DST :	BOOL;
		TIME_ZONE_OFFSET :	INT;
	END_VAR

	LTIME_TO_UTC := LTIME - _INT_TO_UDINT(TIME_ZONE_OFFSET * 60);
	IF DST THEN LTIME_TO_UTC := LTIME_TO_UTC - UDINT#3600; END_IF;

END_FUNCTION

PROGRAM program0
	VAR
		LTIME :	UDINT;
		DST :	BOOL;
		TIME_ZONE_OFFSET :	INT;
		CEIL5_OUT : UDINT;
	END_VAR

  CEIL5_OUT := LTIME_TO_UTC(LTIME, DST, TIME_ZONE_OFFSET);
END_PROGRAM

CONFIGURATION Config0

  RESOURCE Res0 ON PLC
    TASK task0(INTERVAL := T#20ms,PRIORITY := 0);
    PROGRAM instance0 WITH task0 : program0;
  END_RESOURCE
END_CONFIGURATION

(* ---- 25-TRUNC_REAL.ST ---- *)
FUNCTION TRUNC_REAL:REAL

	VAR_INPUT
		IN :	REAL;
	END_VAR

	TRUNC_REAL := UDINT_TO_REAL(DINT_TO_UDINT(TRUNC(IN)));
END_FUNCTION

PROGRAM program0

	VAR
		IN :	REAL;
		OUT: REAL;
	END_VAR
	OUT := TRUNC_REAL(IN);

END_PROGRAM

CONFIGURATION Config0

	RESOURCE Res0 ON PLC
		TASK task0(INTERVAL := T#20ms,PRIORITY := 0);
		PROGRAM instance0 WITH task0 : program0;
	END_RESOURCE

END_CONFIGURATION

(* ---- 252-DEW_CON.ST ---- *)
FUNCTION SDD:REAL

	VAR_INPUT
		T :	REAL;
		ICE :	BOOL;
	END_VAR

	IF ice THEN
		SDD := 611.153 * EXP(22.4433 * T / (272.186 + T));
	ELSE
		SDD := 611.213 * EXP(17.5043 * T / (241.2 + T));
	END_IF;

END_FUNCTION

FUNCTION DEW_CON:REAL

	VAR_INPUT
		RH :	REAL;
		T :	REAL;
	END_VAR

	IF RH > 0.0 AND T > -50.0 THEN
		DEW_CON := 2.166824303E-2 * RH * SDD(T,FALSE)  / (T - -273.15);
	ELSE
		DEW_CON := 0.0;
	END_IF;

END_FUNCTION

PROGRAM program0
  VAR
    RH :	REAL;
	T :	REAL;
    CEIL5_OUT : REAL;
  END_VAR

  CEIL5_OUT := DEW_CON(RH, T);
END_PROGRAM

CONFIGURATION Config0

  RESOURCE Res0 ON PLC
    TASK task0(INTERVAL := T#20ms,PRIORITY := 0);
    PROGRAM instance0 WITH task0 : program0;
  END_RESOURCE
END_CONFIGURATION

(* ---- 254-FIB.ST ---- *)
FUNCTION FIB:DINT

VAR_INPUT
	X :	INT;
END_VAR

VAR
	t1 :	DINT;
	t2 :	DINT;
	X_tmp :	INT;
END_VAR

t1 := DINT#0;
t2 := DINT#0;
X_tmp := X;
IF X_tmp < 0 OR X_tmp > 46 THEN
	FIB := DINT#-1;
ELSIF X_tmp < 2 THEN
	FIB := INT_TO_DINT(X_tmp);
	RETURN;
ELSE
	t2 := DINT#1;
	WHILE X_tmp > 3 DO
		X_tmp := X_tmp - 2;
		t1 := t1 + t2;
		t2 := t1 + t2;
	END_WHILE;
	IF X_tmp > 2 THEN t1 := t1 + t2; END_IF;
	fib := t1 + t2;
END_IF;

END_FUNCTION

PROGRAM program0
  VAR
    LocalVar0 : INT;
	LocalOUT  : DINT;
  END_VAR
  	LocalOUT := FIB(LocalVar0);
END_PROGRAM

CONFIGURATION Config0
  RESOURCE Res0 ON PLC
    TASK task0(INTERVAL := T#20ms,PRIORITY := 0);
    PROGRAM instance0 WITH task0 : program0;
  END_RESOURCE
END_CONFIGURATION

(* ---- 255-AIR_DENSITY.ST ---- *)
FUNCTION SDD:REAL

	VAR_INPUT
		T :	REAL;
		ICE :	BOOL;
	END_VAR

	IF ice THEN
		SDD := 611.153 * EXP(22.4433 * T / (272.186 + T));
	ELSE
		SDD := 611.213 * EXP(17.5043 * T / (241.2 + T));
	END_IF;

END_FUNCTION

FUNCTION AIR_DENSITY:REAL

	VAR_INPUT
		T :	REAL;
		P :	REAL;
		RH :	REAL;
	END_VAR

	AIR_DENSITY := 101325.0 * (1.0 - RH * SDD(T, TRUE) * 3.773319E-3 / P) / (287.05 * ( T - -273.15));

END_FUNCTION

PROGRAM program0
  VAR
    T :	REAL;
	P :	REAL;
	RH :	REAL;
    CEIL5_OUT : REAL;
  END_VAR

  CEIL5_OUT := AIR_DENSITY(T, P, RH);
END_PROGRAM

CONFIGURATION Config0

  RESOURCE Res0 ON PLC
    TASK task0(INTERVAL := T#20ms,PRIORITY := 0);
    PROGRAM instance0 WITH task0 : program0;
  END_RESOURCE
END_CONFIGURATION

(* ---- 256-ISC_ALPHA.ST ---- *)
FUNCTION SETUP_EXTENDED_ASCII:BOOL

	VAR_INPUT
		X :	BOOL;
	END_VAR

	SETUP_EXTENDED_ASCII := X OR TRUE;

END_FUNCTION

FUNCTION ISC_ALPHA:BOOL

	VAR_INPUT
		IN :	BYTE;
	END_VAR

	IF SETUP_EXTENDED_ASCII(FALSE) THEN
		ISC_ALPHA := (in > BYTE#64 AND in < BYTE#91) OR (in > BYTE#191  AND in <> BYTE#215 AND in <> BYTE#247) OR (in > BYTE#96 AND in < BYTE#123);
	ELSE
		ISC_ALPHA := (IN > BYTE#64 AND IN < BYTE#91) OR (in > BYTE#96 AND in < BYTE#123);
	END_IF;

END_FUNCTION

PROGRAM program0
	VAR
		IN : BYTE;
		OUT : BOOL;
	END_VAR

	OUT := ISC_ALPHA(IN);
END_PROGRAM

CONFIGURATION Config0

	RESOURCE Res0 ON PLC
		TASK task0(INTERVAL := T#20ms,PRIORITY := 0);
		PROGRAM instance0 WITH task0 : program0;
	END_RESOURCE

END_CONFIGURATION

(* ---- 259-BINOM.ST ---- *)
FUNCTION BINOM:INT
	VAR_INPUT
		N :	INT;
		K :	INT;
	END_VAR

	VAR
		i :	INT;
		N2 :	INT;
		K2 :	INT;
	END_VAR

	K2 := K;
	N2 := N;
	IF 2 * K2 > N2 THEN
		K2 := N2 - K2;
	END_IF;
	IF K2 > N2 THEN
		RETURN;
	ELSIF K2 = 0 OR K2 = N2 THEN
		BINOM := 1;
	ELSIF K2 = 1 THEN
		BINOM := N2;
	ELSE
		BINOM := N2;
		N2 := N2 + 1;
		FOR i := 2 TO K2 DO
			BINOM := BINOM * (N2 - i) / i;
		END_FOR;
	END_IF;
END_FUNCTION

PROGRAM program0
  VAR
    LocalVar0 : INT;
	LocalVar1 : INT;
    LocalOUT  : INT;
  END_VAR

  LocalOUT := BINOM(LocalVar0, LocalVar1);
END_PROGRAM

CONFIGURATION Config0
  RESOURCE Res0 ON PLC
    TASK task0(INTERVAL := T#20ms,PRIORITY := 0);
    PROGRAM instance0 WITH task0 : program0;
  END_RESOURCE
END_CONFIGURATION

(* ---- 26-ACOTH.ST ---- *)
FUNCTION ACOTH:REAL
	VAR_INPUT
		X :	REAL;
	END_VAR

	ACOTH := LN((x+1.0)/(x-1.0))*0.5;

END_FUNCTION

PROGRAM program0
  VAR
    LocalVar0 : REAL;
    LocalOUT  : REAL;
  END_VAR

  LocalOUT := ACOTH(LocalVar0);
END_PROGRAM

CONFIGURATION Config0
  RESOURCE Res0 ON PLC
    TASK task0(INTERVAL := T#20ms,PRIORITY := 0);
    PROGRAM instance0 WITH task0 : program0;
  END_RESOURCE
END_CONFIGURATION

(* ---- 262-WATER_DENSITY.ST ---- *)
FUNCTION WATER_DENSITY:REAL

    VAR_INPUT
        T :	REAL;
        SAT :	BOOL;
    END_VAR

    VAR
        T2 :	REAL;
        T4 :	REAL;
    END_VAR

    T2 := T * T;
    T4 := T2 * T2;
    WATER_DENSITY := (999.83952 + 16.952577*T + -7.9905127E-3*T2 + -4.6241757E-5*T2*T + 1.0584601E-7*T4 + -2.8103006E-10*T4*T) / (1.0 + 0.0168872*T);
    IF sat THEN WATER_DENSITY := WATER_DENSITY - 0.004612 + 0.000106 * T; END_IF;

END_FUNCTION

PROGRAM program0
	VAR
		T :	REAL;
        SAT :	BOOL;
		CEIL5_OUT : REAL;
	END_VAR

  	CEIL5_OUT := WATER_DENSITY(T, SAT);
END_PROGRAM

CONFIGURATION Config0

  RESOURCE Res0 ON PLC
    TASK task0(INTERVAL := T#20ms,PRIORITY := 0);
    PROGRAM instance0 WITH task0 : program0;
  END_RESOURCE
END_CONFIGURATION

(* ---- 263-FRACT.ST ---- *)
FUNCTION D_TRUNC : DINT
  VAR_INPUT
    x : REAL;
  END_VAR

  D_TRUNC := REAL_TO_DINT(X);
  IF X > 0.0 THEN
  	IF DINT_TO_REAL(D_TRUNC) > X THEN D_TRUNC := D_TRUNC - DINT#1; END_IF;
  ELSE
  	IF DINT_TO_REAL(D_TRUNC) < X THEN D_TRUNC := D_TRUNC + DINT#1; END_IF;
  END_IF;
END_FUNCTION

FUNCTION FRACT:REAL
	VAR_INPUT
		X :	REAL;
	END_VAR

	IF ABS(x) < 2.0E9 THEN
		FRACT := x - DINT_TO_REAL(D_TRUNC(x));
	ELSE
		FRACT := 0.0;
	END_IF;
END_FUNCTION

PROGRAM program0
  VAR
    LocalVar0 : REAL;
	LocalOUT  : REAL;
  END_VAR
  	LocalOUT := FRACT(LocalVar0);
END_PROGRAM

CONFIGURATION Config0
  RESOURCE Res0 ON PLC
    TASK task0(INTERVAL := T#20ms,PRIORITY := 0);
    PROGRAM instance0 WITH task0 : program0;
  END_RESOURCE
END_CONFIGURATION

(* ---- 264-HOUR_TO_TOD.ST ---- *)
FUNCTION _REAL_TO_UDINT:UDINT
	VAR_INPUT
		X :	REAL;
	END_VAR

	IF REAL_TO_UDINT(0.5) = UDINT#1 THEN
		_REAL_TO_UDINT := REAL_TO_UDINT(x);
	ELSIF X > 0.0 THEN
		_REAL_TO_UDINT := REAL_TO_UDINT(x+0.5);
	ELSIF X < 0.0 THEN
		_REAL_TO_UDINT := REAL_TO_UDINT(x-0.5);
	ELSE
		_REAL_TO_UDINT := UDINT#0;
	END_IF;

END_FUNCTION

FUNCTION HOUR_TO_TOD:UDINT

	VAR_INPUT
		IN :	REAL;
	END_VAR

	hour_to_tod := _REAL_TO_UDINT(IN * 3600000.00);

END_FUNCTION

PROGRAM program0
	VAR
		IN :	REAL;
		CEIL5_OUT : UDINT;
	END_VAR

  	CEIL5_OUT := HOUR_TO_TOD(IN);
END_PROGRAM

CONFIGURATION Config0

  RESOURCE Res0 ON PLC
    TASK task0(INTERVAL := T#20ms,PRIORITY := 0);
    PROGRAM instance0 WITH task0 : program0;
  END_RESOURCE

END_CONFIGURATION

(* ---- 267-SCALE_D.ST ---- *)
FUNCTION SCALE_D:REAL
	VAR_INPUT
		X :	DWORD;
		I_LO :	DWORD;
		I_HI :	DWORD;
		O_LO :	REAL;
		O_HI :	REAL;
	END_VAR
	IF I_HI = I_LO THEN
		SCALE_D := O_LO;
	ELSE
		SCALE_D := (O_HI - O_LO) / UDINT_TO_REAL(DWORD_TO_UDINT(I_HI) - DWORD_TO_UDINT(I_LO)) * UDINT_TO_REAL(LIMIT(DWORD_TO_UDINT(I_LO),DWORD_TO_UDINT(X),DWORD_TO_UDINT(I_HI)) - DWORD_TO_UDINT(I_LO)) + O_LO;
	END_IF;
END_FUNCTION

PROGRAM program0
  VAR
		X :	DWORD;
		I_LO :	DWORD;
		I_HI :	DWORD;
		O_LO :	REAL;
		O_HI :	REAL;
		CEIL5_OUT : REAL;
  END_VAR

  CEIL5_OUT := SCALE_D(X, I_LO, I_HI, O_LO, O_HI);
END_PROGRAM

CONFIGURATION Config0

  RESOURCE Res0 ON PLC
    TASK task0(INTERVAL := T#20ms,PRIORITY := 0);
    PROGRAM instance0 WITH task0 : program0;
  END_RESOURCE
END_CONFIGURATION

(* ---- 27-JD2000.ST ---- *)
FUNCTION JD2000:REAL

	VAR_INPUT
		DTI :	UDINT;
	END_VAR

	JD2000 := UDINT_TO_REAL(DTI - UDINT#946728000) / 86400.0;

END_FUNCTION

PROGRAM program0
	VAR
		DTI :	UDINT;
		OUT : REAL;
	END_VAR

	OUT := JD2000(DTI);
END_PROGRAM

CONFIGURATION Config0

	RESOURCE Res0 ON PLC
		TASK task0(INTERVAL := T#20ms,PRIORITY := 0);
		PROGRAM instance0 WITH task0 : program0;
	END_RESOURCE

END_CONFIGURATION

(* ---- 270-HOUR_TO_TIME.ST ---- *)
FUNCTION _REAL_TO_UDINT:UDINT
	VAR_INPUT
		X :	REAL;
	END_VAR

	IF REAL_TO_UDINT(0.5) = UDINT#1 THEN
		_REAL_TO_UDINT := REAL_TO_UDINT(x);
	ELSIF X > 0.0 THEN
		_REAL_TO_UDINT := REAL_TO_UDINT(x+0.5);
	ELSIF X < 0.0 THEN
		_REAL_TO_UDINT := REAL_TO_UDINT(x-0.5);
	ELSE
		_REAL_TO_UDINT := UDINT#0;
  	END_IF;
END_FUNCTION

FUNCTION HOUR_TO_TIME:TIME

	VAR_INPUT
		IN :	REAL;
	END_VAR

	hour_to_time := UDINT_TO_TIME(_REAL_TO_UDINT(IN * 3600000.0));

END_FUNCTION

PROGRAM program0

	VAR
		IN :	REAL;
		CEIL5_OUT : TIME;
	END_VAR

  	CEIL5_OUT := HOUR_TO_TIME(IN);

END_PROGRAM

CONFIGURATION Config0

	RESOURCE Res0 ON PLC
		TASK task0(INTERVAL := T#20ms,PRIORITY := 0);
		PROGRAM instance0 WITH task0 : program0;
	END_RESOURCE

END_CONFIGURATION

(* ---- 272-SECOND_TO_TIME.ST ---- *)
FUNCTION _REAL_TO_UDINT:UDINT
	VAR_INPUT
		X :	REAL;
	END_VAR

	IF REAL_TO_UDINT(0.5) = UDINT#1 THEN
		_REAL_TO_UDINT := REAL_TO_UDINT(x);
	ELSIF X > 0.0 THEN
		_REAL_TO_UDINT := REAL_TO_UDINT(x+0.5);
	ELSIF X < 0.0 THEN
		_REAL_TO_UDINT := REAL_TO_UDINT(x-0.5);
	ELSE
		_REAL_TO_UDINT := UDINT#0;
	END_IF;
END_FUNCTION

FUNCTION SECOND_TO_TIME:TIME

	VAR_INPUT
		IN :	REAL;
	END_VAR

	second_to_time := UDINT_TO_TIME(_REAL_TO_UDINT(IN * 1000.0));

END_FUNCTION

PROGRAM program0

	VAR
		IN :	REAL;
		CEIL5_OUT : TIME;
	END_VAR

	CEIL5_OUT := SECOND_TO_TIME(IN);

END_PROGRAM

CONFIGURATION Config0

	RESOURCE Res0 ON PLC
		TASK task0(INTERVAL := T#20ms,PRIORITY := 0);
		PROGRAM instance0 WITH task0 : program0;
	END_RESOURCE

END_CONFIGURATION

(* ---- 274-MINUTE_TO_TIME.ST ---- *)
FUNCTION _REAL_TO_UDINT:UDINT

  	VAR_INPUT
		X :	REAL;
	END_VAR

	IF REAL_TO_UDINT(0.5) = UDINT#1 THEN
		_REAL_TO_UDINT := REAL_TO_UDINT(x);
	ELSIF X > 0.0 THEN
		_REAL_TO_UDINT := REAL_TO_UDINT(x+0.5);
	ELSIF X < 0.0 THEN
		_REAL_TO_UDINT := REAL_TO_UDINT(x-0.5);
	ELSE
		_REAL_TO_UDINT := UDINT#0;
	END_IF;

END_FUNCTION

FUNCTION MINUTE_TO_TIME:TIME

	VAR_INPUT
		IN :	REAL;
	END_VAR

	minute_to_time := UDINT_TO_TIME(_REAL_TO_UDINT(IN * 60000.0));

END_FUNCTION

PROGRAM program0

	VAR
		IN :	REAL;
		CEIL5_OUT : TIME;
	END_VAR

	CEIL5_OUT := MINUTE_TO_TIME(IN);

END_PROGRAM

CONFIGURATION Config0

	RESOURCE Res0 ON PLC
		TASK task0(INTERVAL := T#20ms,PRIORITY := 0);
		PROGRAM instance0 WITH task0 : program0;
	END_RESOURCE

END_CONFIGURATION

(* ---- 275-F_TO_PT.ST ---- *)
FUNCTION _REAL_TO_DWORD: DWORD
  VAR_INPUT
    X :	REAL;
  END_VAR

  IF REAL_TO_DWORD(0.5) = DWORD#1 THEN
    _REAL_TO_DWORD := REAL_TO_DWORD(x);
  ELSIF X > 0.0 THEN
    _REAL_TO_DWORD := REAL_TO_DWORD(x+0.5);
  ELSIF X < 0.0 THEN
    _REAL_TO_DWORD := REAL_TO_DWORD(x-0.5);
  ELSE
    _REAL_TO_DWORD := DWORD#0;
  END_IF;
END_FUNCTION

FUNCTION F_TO_PT:TIME
	VAR_INPUT
		F :	REAL;
	END_VAR
	F_TO_PT := DWORD_TO_TIME(_REAL_TO_DWORD(1.0 / F * 1000.0));
END_FUNCTION

PROGRAM program0
  VAR
    LocalVar0 : REAL;
	  LocalOUT  : TIME;
  END_VAR
  	LocalOUT := F_TO_PT(LocalVar0);
END_PROGRAM

CONFIGURATION Config0
  RESOURCE Res0 ON PLC
    TASK task0(INTERVAL := T#20ms,PRIORITY := 0);
    PROGRAM instance0 WITH task0 : program0;
  END_RESOURCE
END_CONFIGURATION

(* ---- 276-ATAN2.ST ---- *)
FUNCTION ATAN2:REAL
	VAR_INPUT
		X :	REAL;
		Y :	REAL;
	END_VAR

	IF X > 0.0 THEN
		ATAN2 := ATAN(Y/X);
	ELSIF X < 0.0 THEN
		IF Y >= 0.0 THEN
			ATAN2 := ATAN(Y/X) + 3.14159265358979323846264338327950288;
		ELSE
			ATAN2 := ATAN(Y/X) - 3.14159265358979323846264338327950288;
		END_IF;
	ELSIF Y > 0.0 THEN
		ATAN2 := 1.5707963267948965580;
	ELSIF Y < 0.0 THEN
		ATAN2 := -1.5707963267948965580;
	ELSE
		ATAN2 := 0.0;
	END_IF;

END_FUNCTION

PROGRAM program0
  VAR
    LocalVar0 : REAL;
	LocalVar1 : REAL;
    LocalOUT  : REAL;
  END_VAR

  LocalOUT := ATAN2(LocalVar0, LocalVar1);
END_PROGRAM

CONFIGURATION Config0
  RESOURCE Res0 ON PLC
    TASK task0(INTERVAL := T#20ms,PRIORITY := 0);
    PROGRAM instance0 WITH task0 : program0;
  END_RESOURCE
END_CONFIGURATION

(* ---- 277-DEG.ST ---- *)
FUNCTION FLOOR2 : DINT
	VAR_INPUT
		x : REAL;
	END_VAR

	FLOOR2 := REAL_TO_DINT(X);
	IF DINT_TO_REAL(FLOOR2) > X THEN
		FLOOR2 := FLOOR2 - DINT#1;
	END_IF;

END_FUNCTION

FUNCTION MODR:REAL

	VAR_INPUT
		IN :	REAL;
		DIVI :	REAL;
	END_VAR

	IF divi = 0.0 THEN
		MODR := 0.0;
	ELSE
		MODR := in - DINT_TO_REAL(FLOOR2(in / divi)) * divi;
	END_IF;

END_FUNCTION

FUNCTION DEG:REAL

	VAR_INPUT
		RAD :	REAL;
	END_VAR

	DEG := MODR(57.29577951308232 * RAD, 360.0);

END_FUNCTION

PROGRAM program0

	VAR
		RAD :	REAL;
		CEIL5_OUT : REAL;
	END_VAR

	CEIL5_OUT := DEG(RAD);

END_PROGRAM

CONFIGURATION Config0

	RESOURCE Res0 ON PLC
		TASK task0(INTERVAL := T#20ms,PRIORITY := 0);
		PROGRAM instance0 WITH task0 : program0;
	END_RESOURCE

END_CONFIGURATION

(* ---- 28-SIGN_R.ST ---- *)
FUNCTION SIGN_R : BOOL
  VAR_INPUT
    IN : REAL;
  END_VAR

  SIGN_R := in < 0.0;
END_FUNCTION

PROGRAM program0
  VAR
    LocalVar0 : REAL;
    CEIL5_OUT : BOOL;
  END_VAR

  CEIL5_OUT := SIGN_R(LocalVar0);
END_PROGRAM

CONFIGURATION Config0

  RESOURCE Res0 ON PLC
    TASK task0(INTERVAL := T#20ms,PRIORITY := 0);
    PROGRAM instance0 WITH task0 : program0;
  END_RESOURCE
END_CONFIGURATION

(* ---- 285-BYTE_OF_BIT.ST ---- *)
FUNCTION BYTE_OF_BIT:BYTE
	VAR_INPUT
		B0 :	BOOL;
		B1 :	BOOL;
		B2 :	BOOL;
		B3 :	BOOL;
		B4 :	BOOL;
		B5 :	BOOL;
		B6 :	BOOL;
		B7 :	BOOL;
	END_VAR
	Byte_of_bit := SHL(SHL(SHL(SHL(SHL(SHL(SHL(BOOL_TO_BYTE(B7),1) OR BOOL_TO_BYTE(B6),1)
	OR BOOL_TO_BYTE(B5),1) OR BOOL_TO_BYTE(B4),1) OR BOOL_TO_BYTE(B3),1) OR BOOL_TO_BYTE(B2),1)
	OR BOOL_TO_BYTE(B1),1) OR BOOL_TO_BYTE(B0);
END_FUNCTION

PROGRAM program0
  VAR
	B0 :	BOOL;
	B1 :	BOOL;
	B2 :	BOOL;
	B3 :	BOOL;
	B4 :	BOOL;
	B5 :	BOOL;
	B6 :	BOOL;
	B7 :	BOOL;
    LocalOUT  : BYTE;
  END_VAR

  LocalOUT := BYTE_OF_BIT(B0, B1, B2, B3, B4, B5, B6, B7);
END_PROGRAM

CONFIGURATION Config0
  RESOURCE Res0 ON PLC
    TASK task0(INTERVAL := T#20ms,PRIORITY := 0);
    PROGRAM instance0 WITH task0 : program0;
  END_RESOURCE
END_CONFIGURATION

(* ---- 286-RAD.ST ---- *)
FUNCTION FLOOR2 : DINT
	VAR_INPUT
		x : REAL;
	END_VAR

	FLOOR2 := REAL_TO_DINT(X);
	IF DINT_TO_REAL(FLOOR2) > X THEN
		FLOOR2 := FLOOR2 - DINT#1;
	END_IF;

END_FUNCTION

FUNCTION MODR: REAL

	VAR_INPUT
		IN :	REAL;
		DIVI :	REAL;
	END_VAR

	IF divi = 0.0 THEN
		MODR := 0.0;
	ELSE
		MODR := in - DINT_TO_REAL(FLOOR2(in / divi)) * divi;
	END_IF;

END_FUNCTION

FUNCTION RAD:REAL

	VAR_INPUT
		DEG :	REAL;
	END_VAR

	RAD := MODR(0.0174532925199433 * DEG , 6.283185307179586476);

END_FUNCTION

PROGRAM program0

	VAR
		DEG :	REAL;
		CEIL5_OUT : REAL;
	END_VAR

	CEIL5_OUT := RAD(DEG);

END_PROGRAM

CONFIGURATION Config0

	RESOURCE Res0 ON PLC
		TASK task0(INTERVAL := T#20ms,PRIORITY := 0);
		PROGRAM instance0 WITH task0 : program0;
	END_RESOURCE

END_CONFIGURATION

(* ---- 287-REAL_TO_TIME.ST ---- *)
FUNCTION _REAL_TO_UDINT:UDINT
  VAR_INPUT
    X :	REAL;
  END_VAR

  IF REAL_TO_UDINT(0.5) = UDINT#1 THEN
    _REAL_TO_UDINT := REAL_TO_UDINT(x);
  ELSIF X > 0.0 THEN
    _REAL_TO_UDINT := REAL_TO_UDINT(x+0.5);
  ELSIF X < 0.0 THEN
    _REAL_TO_UDINT := REAL_TO_UDINT(x-0.5);
  ELSE
    _REAL_TO_UDINT := UDINT#0;
  END_IF;
END_FUNCTION

FUNCTION REAL_TO_TIME2:TIME
	VAR_INPUT
		IN :	REAL;
	END_VAR

	REAL_TO_TIME2 := DINT_TO_TIME(UDINT_TO_DINT(_REAL_TO_UDINT(IN)));
END_FUNCTION

PROGRAM program0
  VAR
    LocalVar0 : REAL;
    LocalOUT  : TIME;
  END_VAR

  LocalOUT := REAL_TO_TIME2(LocalVar0);
END_PROGRAM

CONFIGURATION Config0
  RESOURCE Res0 ON PLC
    TASK task0(INTERVAL := T#20ms,PRIORITY := 0);
    PROGRAM instance0 WITH task0 : program0;
  END_RESOURCE
END_CONFIGURATION

(* ---- 289-DAY_TO_TIME.ST ---- *)
FUNCTION DAY_TO_TIME:TIME
	VAR_INPUT
		IN :	REAL;
	END_VAR

	day_to_time := DINT_TO_TIME(UDINT_TO_DINT(_REAL_TO_UDINT(IN * REAL#86400000.00)));
END_FUNCTION

FUNCTION _REAL_TO_UDINT:UDINT
  VAR_INPUT
    X :	REAL;
  END_VAR

  IF REAL_TO_UDINT(0.5) = UDINT#1 THEN
    _REAL_TO_UDINT := REAL_TO_UDINT(x);
  ELSIF X > 0.0 THEN
    _REAL_TO_UDINT := REAL_TO_UDINT(x+0.5);
  ELSIF X < 0.0 THEN
    _REAL_TO_UDINT := REAL_TO_UDINT(x-0.5);
  ELSE
    _REAL_TO_UDINT := UDINT#0;
  END_IF;
END_FUNCTION

PROGRAM program0
  VAR
    LocalVar0 : REAL;
	LocalOUT  : TIME;
  END_VAR
  	LocalOUT := DAY_TO_TIME(LocalVar0);
END_PROGRAM

CONFIGURATION Config0
  RESOURCE Res0 ON PLC
    TASK task0(INTERVAL := T#20ms,PRIORITY := 0);
    PROGRAM instance0 WITH task0 : program0;
  END_RESOURCE
END_CONFIGURATION

(* ---- 29-TRUNC_UDINT.ST ---- *)
FUNCTION TRUNC_UDINT:UDINT
	VAR_INPUT
		IN :	REAL;
	END_VAR
	TRUNC_UDINT := DINT_TO_UDINT(TRUNC(IN));
END_FUNCTION

PROGRAM program0
	VAR
		LocalVar0 : REAL;
		LocalOUT  : UDINT;
	END_VAR
		LocalOUT := TRUNC_UDINT(LocalVar0);
END_PROGRAM

CONFIGURATION Config0
	RESOURCE Res0 ON PLC
		TASK task0(INTERVAL := T#20ms,PRIORITY := 0);
		PROGRAM instance0 WITH task0 : program0;
	END_RESOURCE
END_CONFIGURATION

(* ---- 290-ERFC.ST ---- *)
FUNCTION SGN : INT
  VAR_INPUT
    x : REAL;
  END_VAR

  IF X > 0.0 THEN
  	sgn := 1;
  ELSIF X < 0.0 THEN
  	sgn := -1;
  ELSE
  	sgn := 0;
  END_IF;
END_FUNCTION

FUNCTION ERF:REAL

	VAR_INPUT
		X :	REAL;
	END_VAR

	VAR
		x2 :	REAL;
		ax2 :	REAL;
	END_VAR

	x2 := X*X;
	ax2 := 0.147 * x2 + 1.0;
	ERF := SQRT(1.0 - EXP(-X2 * ((0.27323954473516 + aX2)/(ax2)))) * INT_TO_REAL(SGN(x));

END_FUNCTION

FUNCTION ERFC:REAL
	VAR_INPUT
		X :	REAL;
	END_VAR

	ERFC := 1.0 - ERF(X);

END_FUNCTION

PROGRAM program0
  VAR
    LocalVar0 : REAL;
	  LocalOUT  : REAL;
  END_VAR
  	LocalOUT := ERFC(LocalVar0);
END_PROGRAM

CONFIGURATION Config0
  RESOURCE Res0 ON PLC
    TASK task0(INTERVAL := T#20ms,PRIORITY := 0);
    PROGRAM instance0 WITH task0 : program0;
  END_RESOURCE
END_CONFIGURATION

(* ---- 293-SCALE_B.ST ---- *)
FUNCTION _BYTE_TO_REAL:REAL
	VAR_INPUT
		IN :	BYTE;
	END_VAR

	_BYTE_TO_REAL := USINT_TO_REAL(BYTE_TO_USINT(IN));
END_FUNCTION

FUNCTION SCALE_B:REAL

	VAR_INPUT
		X :	BYTE;
		I_LO :	BYTE;
		I_HI :	BYTE;
		O_LO :	REAL;
		O_HI :	REAL;
	END_VAR

	IF I_HI = I_LO THEN
		SCALE_B := O_LO;
	ELSE
		SCALE_B := (O_HI - O_LO) / USINT_TO_REAL(BYTE_TO_USINT(I_HI) - BYTE_TO_USINT(I_LO)) * _BYTE_TO_REAL(LIMIT(I_LO,X,I_HI));
	END_IF;

END_FUNCTION

PROGRAM program0
  VAR
	X :	BYTE;
	I_LO :	BYTE;
	I_HI :	BYTE;
	O_LO :	REAL;
	O_HI :	REAL;
	CEIL5_OUT : REAL;
  END_VAR

  CEIL5_OUT := SCALE_B(X, I_LO, I_HI, O_LO, O_HI);

END_PROGRAM

CONFIGURATION Config0

  RESOURCE Res0 ON PLC
    TASK task0(INTERVAL := T#20ms,PRIORITY := 0);
    PROGRAM instance0 WITH task0 : program0;
  END_RESOURCE
END_CONFIGURATION

(* ---- 295-STAIR.ST ---- *)
FUNCTION _REAL_TO_DINT:DINT
	VAR_INPUT
		X :	REAL;
	END_VAR

	IF REAL_TO_DINT(0.5) = DINT#1 THEN
		_REAL_TO_DINT := REAL_TO_DINT(x);
		RETURN;
	END_IF;

	IF X > 0.0 THEN
		_REAL_TO_DINT := REAL_TO_DINT(x+0.5);
	ELSIF X < 0.0 THEN
		_REAL_TO_DINT := REAL_TO_DINT(x-0.5);
	ELSE
		_REAL_TO_DINT := DINT#0;
	END_IF;

END_FUNCTION

FUNCTION STAIR:REAL

	VAR_INPUT
		X :	REAL;
		D :	REAL;
	END_VAR

	IF D > 0.0 THEN
		STAIR := DINT_TO_REAL(_REAL_TO_DINT(X / D)) * D;
	ELSE
		STAIR := X;
	END_IF;

END_FUNCTION

PROGRAM program0

	VAR
		X :	REAL;
		D :	REAL;
		CEIL5_OUT : REAL;
	END_VAR

	CEIL5_OUT := STAIR(X, D);

END_PROGRAM

CONFIGURATION Config0

	RESOURCE Res0 ON PLC
		TASK task0(INTERVAL := T#20ms,PRIORITY := 0);
		PROGRAM instance0 WITH task0 : program0;
	END_RESOURCE

END_CONFIGURATION

(* ---- 297-CEIL2.ST ---- *)
FUNCTION _REAL_TO_DINT:DINT
  VAR_INPUT
    X :	REAL;
  END_VAR

  IF REAL_TO_DINT(0.5) = DINT#1 THEN
    _REAL_TO_DINT := REAL_TO_DINT(x);
    RETURN;
  END_IF;

  IF X > 0.0 THEN
    _REAL_TO_DINT := REAL_TO_DINT(x+0.5);
  ELSIF X < 0.0 THEN
    _REAL_TO_DINT := REAL_TO_DINT(x-0.5);
  ELSE
    _REAL_TO_DINT := DINT#0;
  END_IF;
END_FUNCTION

FUNCTION CEIL2:DINT

	VAR_INPUT
		X :	REAL;
	END_VAR

	CEIL2 := _REAL_TO_DINT(x);
	IF DINT_TO_REAL(CEIL2) < X THEN
			CEIL2 := CEIL2 + DINT#1;
	END_IF;

END_FUNCTION

PROGRAM program0
  VAR
    LocalVar0 : REAL;
    CEIL5_OUT : DINT;
  END_VAR

  CEIL5_OUT := CEIL2(LocalVar0);
END_PROGRAM

CONFIGURATION Config0

  RESOURCE Res0 ON PLC
    TASK task0(INTERVAL := T#20ms,PRIORITY := 0);
    PROGRAM instance0 WITH task0 : program0;
  END_RESOURCE
END_CONFIGURATION

(* ---- 30-C_TO_K.ST ---- *)
FUNCTION C_TO_K:REAL
	VAR_INPUT
		CELSIUS :	REAL;
	END_VAR

	C_to_K := Celsius - 273.15;
END_FUNCTION

PROGRAM program0
  VAR
    LocalVar0 : REAL;
    CEIL5_OUT : REAL;
  END_VAR

  CEIL5_OUT := C_TO_K(LocalVar0);
END_PROGRAM

CONFIGURATION Config0

  RESOURCE Res0 ON PLC
    TASK task0(INTERVAL := T#20ms,PRIORITY := 0);
    PROGRAM instance0 WITH task0 : program0;
  END_RESOURCE
END_CONFIGURATION

(* ---- 300-FLOOR2.ST ---- *)
FUNCTION _REAL_TO_DINT:DINT
  VAR_INPUT
    X :	REAL;
  END_VAR

  IF REAL_TO_DINT(0.5) = DINT#1 THEN
    _REAL_TO_DINT := REAL_TO_DINT(x);
    RETURN;
  END_IF;

  IF X > 0.0 THEN
    _REAL_TO_DINT := REAL_TO_DINT(x+0.5);
  ELSIF X < 0.0 THEN
    _REAL_TO_DINT := REAL_TO_DINT(x-0.5);
  ELSE
    _REAL_TO_DINT := DINT#0;
  END_IF;
END_FUNCTION

FUNCTION FLOOR2:DINT
	VAR_INPUT
		X :	REAL;
	END_VAR

	FLOOR2 := _REAL_TO_DINT(X);
	IF DINT_TO_REAL(FLOOR2) > X THEN
		FLOOR2 := FLOOR2 - DINT#1;
	END_IF;
END_FUNCTION

PROGRAM program0
  VAR
    LocalVar0 : REAL;
    CEIL5_OUT : DINT;
  END_VAR

  CEIL5_OUT := FLOOR2(LocalVar0);
END_PROGRAM

CONFIGURATION Config0

  RESOURCE Res0 ON PLC
    TASK task0(INTERVAL := T#20ms,PRIORITY := 0);
    PROGRAM instance0 WITH task0 : program0;
  END_RESOURCE
END_CONFIGURATION

(* ---- 301-CHECK_PARITY.ST ---- *)
FUNCTION BIT_OF_DWORD : BOOL
  VAR_INPUT
    IN : DWORD;
    N : INT;
  END_VAR

  BIT_OF_DWORD := (SHR(in,N) AND 16#00000001) > 0;
END_FUNCTION

FUNCTION CHECK_PARITY:BOOL

	VAR_INPUT
		IN :	DWORD;
		P :	BOOL;
	END_VAR

	VAR
		in2 :	DWORD;
	END_VAR

	in2:=in;
	check_parity := NOT p;
	WHILE in2 > DWORD#0 DO
		check_parity := check_parity XOR BIT_OF_DWORD(in2,0) XOR BIT_OF_DWORD(in2,1) XOR BIT_OF_DWORD(in2,2) XOR BIT_OF_DWORD(in2,3);
		in2 := SHR(in2,4);
	END_WHILE;

END_FUNCTION

PROGRAM program0
  VAR
    LocalVar0 : DWORD;
    LocalVar1 : BOOL;
    CEIL5_OUT : BOOL;
  END_VAR

  CEIL5_OUT := CHECK_PARITY(LocalVar0, LocalVar1);
END_PROGRAM

CONFIGURATION Config0

  RESOURCE Res0 ON PLC
    TASK task0(INTERVAL := T#20ms,PRIORITY := 0);
    PROGRAM instance0 WITH task0 : program0;
  END_RESOURCE
END_CONFIGURATION

(* ---- 304-SCALE_X2.ST ---- *)
FUNCTION SCALE_X2:REAL
	VAR_INPUT
		IN1 :	BOOL;
		IN2 :	BOOL;
		K :	REAL;
		O :	REAL;
		IN1_MIN :	REAL;(*Standard = 0*)
		IN1_MAX :	REAL;(*Standard = 1000*)
		IN2_MIN :	REAL;(*Standard = 0*)
		IN2_MAX :	REAL;(*Standard = 1000*)
	END_VAR

	SCALE_X2 := (SEL(IN1,IN1_MIN, IN1_MAX)+ SEL(IN2,IN2_MIN, IN2_MAX))* k + o;

END_FUNCTION

PROGRAM program0

  	VAR
		IN1 :	BOOL;
		IN2 :	BOOL;
		K :	REAL;
		O :	REAL;
		IN1_MIN :	REAL;(*Standard = 0*)
		IN1_MAX :	REAL;(*Standard = 1000*)
		IN2_MIN :	REAL;(*Standard = 0*)
		IN2_MAX :	REAL;(*Standard = 1000*)
		CEIL5_OUT : REAL;
  	END_VAR

  	CEIL5_OUT := SCALE_X2(IN1, IN2, K, O, IN1_MIN, IN1_MAX, IN2_MIN, IN2_MAX);
END_PROGRAM

CONFIGURATION Config0

	RESOURCE Res0 ON PLC
		TASK task0(INTERVAL := T#20ms,PRIORITY := 0);
		PROGRAM instance0 WITH task0 : program0;
	END_RESOURCE

END_CONFIGURATION

(* ---- 31-MS_TO_BFT.ST ---- *)
FUNCTION MS_TO_BFT:INT

	VAR_INPUT
		MS :	REAL;
	END_VAR

	MS_TO_BFT := REAL_TO_INT(EXPT(MS * 1.196172, 0.666667));

END_FUNCTION

PROGRAM program0
	VAR
		MS :	REAL;

		OUT : INT;
	END_VAR

	OUT := MS_TO_BFT(MS);

END_PROGRAM

CONFIGURATION Config0

	RESOURCE Res0 ON PLC
		TASK task0(INTERVAL := T#20ms,PRIORITY := 0);
		PROGRAM instance0 WITH task0 : program0;
	END_RESOURCE

END_CONFIGURATION

(* ---- 317-DEW_RH.ST ---- *)
FUNCTION SDD:REAL

	VAR_INPUT
		T :	REAL;
		ICE :	BOOL;
	END_VAR

	IF ice THEN
		SDD := 611.153 * EXP(22.4433 * T / (272.186 + T));
	ELSE
		SDD := 611.213 * EXP(17.5043 * T / (241.2 + T));
	END_IF;

END_FUNCTION

FUNCTION DEW_CON:REAL

	VAR_INPUT
		RH :	REAL;
		T :	REAL;
	END_VAR

	IF RH > 0.0 AND T > -50.0 THEN
		DEW_CON := 2.166824303E-2 * RH * SDD(T,FALSE)  / (T - -273.15);
	ELSE
		DEW_CON := 0.0;
	END_IF;

END_FUNCTION

FUNCTION DEW_RH:REAL

	VAR_INPUT
		VC :	REAL;
		T :	REAL;
	END_VAR

	DEW_RH := LIMIT(0.0, VC / DEW_CON(1.0, T), 100.0);

END_FUNCTION

PROGRAM program0
	VAR
		VC :	REAL;
		T :	REAL;
		CEIL5_OUT : REAL;
	END_VAR

  	CEIL5_OUT := DEW_RH(VC, T);
END_PROGRAM

CONFIGURATION Config0

  RESOURCE Res0 ON PLC
    TASK task0(INTERVAL := T#20ms,PRIORITY := 0);
    PROGRAM instance0 WITH task0 : program0;
  END_RESOURCE
END_CONFIGURATION

(* ---- 32-ATANH.ST ---- *)
FUNCTION ATANH:REAL
	VAR_INPUT
		X :	REAL;
	END_VAR

	ATANH := LN((1.0 + x)/(1.0 - x)) * 0.5;

END_FUNCTION

PROGRAM program0
  VAR
    LocalVar0 : REAL;
    LocalOUT  : REAL;
  END_VAR

  LocalOUT := ATANH(LocalVar0);
END_PROGRAM

CONFIGURATION Config0
  RESOURCE Res0 ON PLC
    TASK task0(INTERVAL := T#20ms,PRIORITY := 0);
    PROGRAM instance0 WITH task0 : program0;
  END_RESOURCE
END_CONFIGURATION

(* ---- 324-GAUSSCD.ST ---- *)
FUNCTION SGN : INT
  VAR_INPUT
    x : REAL;
  END_VAR

  IF X > 0.0 THEN
  	sgn := 1;
  ELSIF X < 0.0 THEN
  	sgn := -1;
  ELSE
  	sgn := 0;
  END_IF;
END_FUNCTION

FUNCTION ERF:REAL

	VAR_INPUT
		X :	REAL;
	END_VAR

	VAR
		x2 :	REAL;
		ax2 :	REAL;
	END_VAR

	x2 := X*X;
	ax2 := 0.147 * x2 + 1.0;
	ERF := SQRT(1.0 - EXP(-X2 * ((0.27323954473516 + aX2)/(ax2)))) * INT_TO_REAL(SGN(x));

END_FUNCTION

FUNCTION GAUSSCD:REAL

	VAR_INPUT
		X :	REAL;
		U :	REAL;
		SI :	REAL;
	END_VAR

	GAUSSCD := (ERF((X - U) / (SI * 1.414213562)) + 1.0) * 0.5;

END_FUNCTION

PROGRAM program0
  VAR
    X :	REAL;
	U :	REAL;
	SI :	REAL;
    LocalOUT  : REAL;
  END_VAR

  LocalOUT := GAUSSCD(X, U, SI);
END_PROGRAM

CONFIGURATION Config0
  RESOURCE Res0 ON PLC
    TASK task0(INTERVAL := T#20ms,PRIORITY := 0);
    PROGRAM instance0 WITH task0 : program0;
  END_RESOURCE
END_CONFIGURATION

(* ---- 33-F_TO_OM.ST ---- *)
FUNCTION F_TO_OM:REAL

	VAR_INPUT
		F :	REAL;
	END_VAR

	F_to_OM := 6.283185307179586476 * F;

END_FUNCTION

PROGRAM program0
  VAR
    LocalVar0 : REAL;
	  LocalOUT  : REAL;
  END_VAR
  	LocalOUT := F_TO_OM(LocalVar0);
END_PROGRAM

CONFIGURATION Config0
  RESOURCE Res0 ON PLC
    TASK task0(INTERVAL := T#20ms,PRIORITY := 0);
    PROGRAM instance0 WITH task0 : program0;
  END_RESOURCE
END_CONFIGURATION
